// TIA Portal V19 export
FUNCTION_BLOCK "ALL_PUMPS"   // FB2, LAD
{ S7_Optimized_Access := 'TRUE' }
// stored: MemoryReserve 100, SetENOAutomatically false
   VAR
      PUMP_FB1_CP01 { S7_SetPoint := 'True'} : "PUMP_FB1";
      PUMP_FB1_AG01 { S7_SetPoint := 'True'} : "PUMP_FB1";
      PUMP_FB1_CHS_CP01 { S7_SetPoint := 'True'} : "PUMP_FB1";
      PUMP_FB1_CHS_CP02 { S7_SetPoint := 'True'} : "PUMP_FB1";
      PUMP_FB1_CHS_CP03 { S7_SetPoint := 'True'} : "PUMP_FB1";
      PUMP_FB1_R2_CP01 { S7_SetPoint := 'True'} : "PUMP_FB1";
      PUMP_FB1_R2_AG01 { S7_SetPoint := 'True'} : "PUMP_FB1";
      PUMP_FB1_R3_CP01 { S7_SetPoint := 'True'} : "PUMP_FB1";
      PUMP_FB1_R3_AG01 { S7_SetPoint := 'True'} : "PUMP_FB1";
      PUMP_FB1_R4_CP01 { S7_SetPoint := 'True'} : "PUMP_FB1";
      PUMP_FB1_R4_AG01 { S7_SetPoint := 'True'} : "PUMP_FB1";
      PUMP_FB1_R5_CP01 { S7_SetPoint := 'True'} : "PUMP_FB1";
      PUMP_FB1_R5_AG01 { S7_SetPoint := 'True'} : "PUMP_FB1";
      PUMP_FB1_R6_CP01 { S7_SetPoint := 'True'} : "PUMP_FB1";
      PUMP_FB1_R6_AG01 { S7_SetPoint := 'True'} : "PUMP_FB1";
      PUMP_FB1_R7_CP01 { S7_SetPoint := 'True'} : "PUMP_FB1";
      PUMP_FB1_R7_AG01 { S7_SetPoint := 'True'} : "PUMP_FB1";
      PUMP_FB1_R8_CP01 { S7_SetPoint := 'True'} : "PUMP_FB1";
      PUMP_FB1_R8_AG01 { S7_SetPoint := 'True'} : "PUMP_FB1";
      PUMP_FB1_R9_CP01 { S7_SetPoint := 'True'} : "PUMP_FB1";
      PUMP_FB1_R9_AG01 { S7_SetPoint := 'True'} : "PUMP_FB1";
      PUMP_FB1_R10_CP01 { S7_SetPoint := 'True'} : "PUMP_FB1";
      PUMP_FB1_R10_AG01 { S7_SetPoint := 'True'} : "PUMP_FB1";
      PUMP_FB1_R11_CP01 { S7_SetPoint := 'True'} : "PUMP_FB1";
      PUMP_FB1_R11_AG01 { S7_SetPoint := 'True'} : "PUMP_FB1";
      PUMP_FB1_R12_CP01 { S7_SetPoint := 'True'} : "PUMP_FB1";
      PUMP_FB1_R12_AG01 { S7_SetPoint := 'True'} : "PUMP_FB1";
      PUMP_FB1_R13_CP01 { S7_SetPoint := 'True'} : "PUMP_FB1";
      PUMP_FB1_R13_AG01 { S7_SetPoint := 'True'} : "PUMP_FB1";
      PUMP_FB1_R14_CP01 { S7_SetPoint := 'True'} : "PUMP_FB1";
      PUMP_FB1_R14_AG01 { S7_SetPoint := 'True'} : "PUMP_FB1";
      PUMP_FB1_R15_CP01 { S7_SetPoint := 'True'} : "PUMP_FB1";
      PUMP_FB1_R15_AG01 { S7_SetPoint := 'True'} : "PUMP_FB1";
      PUMP_FB1_R16_CP01 { S7_SetPoint := 'True'} : "PUMP_FB1";
      PUMP_FB1_R16_AG01 { S7_SetPoint := 'True'} : "PUMP_FB1";
      PUMP_FB1_R17_CP01 { S7_SetPoint := 'True'} : "PUMP_FB1";
      PUMP_FB1_R17_AG01 { S7_SetPoint := 'True'} : "PUMP_FB1";
      PUMP_FB1_R18_CP01 { S7_SetPoint := 'True'} : "PUMP_FB1";
      PUMP_FB1_R18_AG01 { S7_SetPoint := 'True'} : "PUMP_FB1";
      PUMP_FB1_CS_CP01 { S7_SetPoint := 'True'} : "PUMP_FB1";
      PUMP_FB1_CS_CP02 { S7_SetPoint := 'True'} : "PUMP_FB1";
      PUMP_FB1_CS_CP03 { S7_SetPoint := 'True'} : "PUMP_FB1";
      PUMP_FB1_UCHS_CP01 { S7_SetPoint := 'True'} : "PUMP_FB1";
      PUMP_FB1_UCHS_CP02 { S7_SetPoint := 'True'} : "PUMP_FB1";
      PUMP_FB1_UCHS_CP03 { S7_SetPoint := 'True'} : "PUMP_FB1";
      PUMP_FB1_HS_CP01 { S7_SetPoint := 'True'} : "PUMP_FB1";
      PUMP_FB1_HS_CP02 { S7_SetPoint := 'True'} : "PUMP_FB1";
      PUMP_FB1_HS_CP03 { S7_SetPoint := 'True'} : "PUMP_FB1";
      "PUMP_FB1_A/SCRB_001_CP01" { S7_SetPoint := 'True'} : "PUMP_FB1";
      "PUMP_FB1_A/SCRB_001_CP02" { S7_SetPoint := 'True'} : "PUMP_FB1";
      "PUMP_FB1_A/SCRB_002_CP01" { S7_SetPoint := 'True'} : "PUMP_FB1";
      "PUMP_FB1_A/SCRB_001_BL01" { S7_SetPoint := 'True'} : "PUMP_FB1";
      "PUMP_FB1_A/SCRB_002_BL02" { S7_SetPoint := 'True'} : "PUMP_FB1";
      "PUMP_FB1_AA/VP_01_CP01" { S7_SetPoint := 'True'} : "PUMP_FB1";
      "PUMP_FB1_A/VP_01_CP01" { S7_SetPoint := 'True'} : "PUMP_FB1";
   END_VAR
BEGIN

REGION Network 1: ***R1****
END_REGION

REGION Network 2: CP01
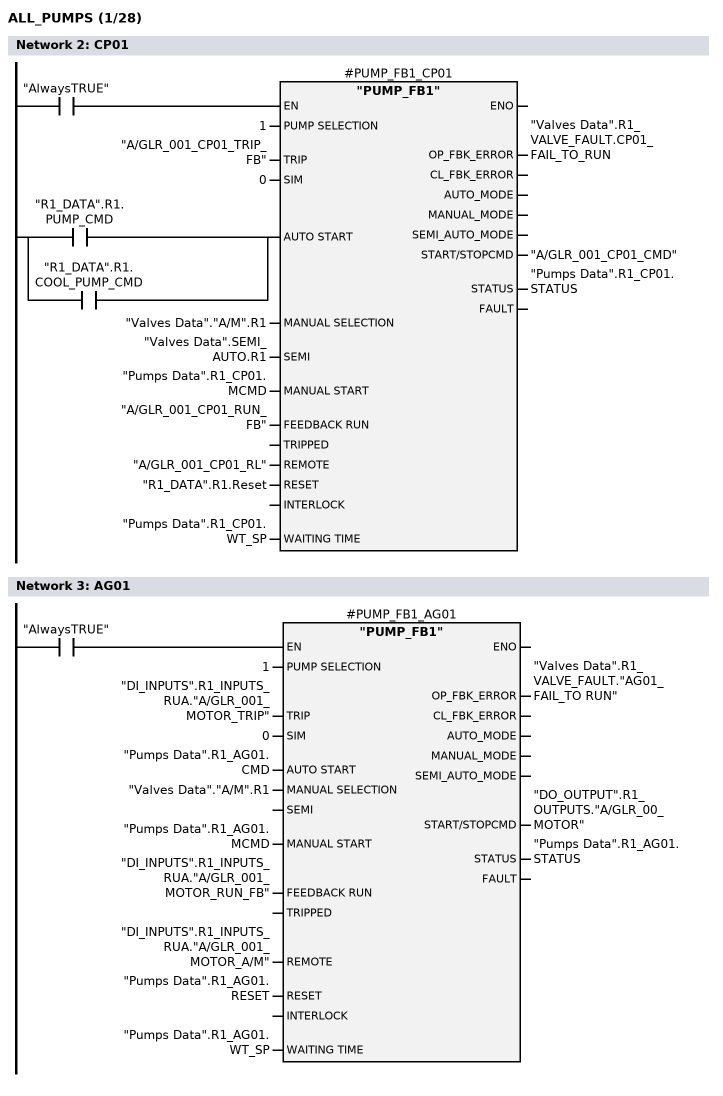
   RUNG wire#powerrail
      Contact( "AlwaysTRUE" )
      #PUMP_FB1_CP01("AUTO START" := wire#w1, "PUMP SELECTION" := 1, TRIP := "A/GLR_001_CP01_TRIP_FB", SIM := 0, "MANUAL SELECTION" := "Valves Data"."A/M".R1, SEMI := "Valves Data".SEMI_AUTO.R1, "MANUAL START" := "Pumps Data".R1_CP01.MCMD, "FEEDBACK RUN" := "A/GLR_001_CP01_RUN_FB", TRIPPED :=, REMOTE := "A/GLR_001_CP01_RL", RESET := "R1_DATA".R1.Reset, INTERLOCK :=, "WAITING TIME" := "Pumps Data".R1_CP01.WT_SP, OP_FBK_ERROR => "Valves Data".R1_VALVE_FAULT.CP01_FAIL_TO_RUN, CL_FBK_ERROR =>, AUTO_MODE =>, MANUAL_MODE =>, SEMI_AUTO_MODE =>, "START/STOPCMD" => "A/GLR_001_CP01_CMD", STATUS => "Pumps Data".R1_CP01.STATUS, FAULT =>)
   END_RUNG
   RUNG wire#powerrail
      Contact( "R1_DATA".R1.PUMP_CMD )
   END_RUNG wire#w1
   RUNG wire#powerrail
      Contact( "R1_DATA".R1.COOL_PUMP_CMD )
   END_RUNG wire#w1
   // the same network as SCL:
   IF "AlwaysTRUE" THEN
       #PUMP_FB1_CP01("PUMP SELECTION" := 1,   // "PUMP_FB1"
                      TRIP := "A/GLR_001_CP01_TRIP_FB",
                      SIM := 0,
                      "AUTO START" := "R1_DATA".R1.PUMP_CMD OR "R1_DATA".R1.COOL_PUMP_CMD,
                      "MANUAL SELECTION" := "Valves Data"."A/M".R1,
                      SEMI := "Valves Data".SEMI_AUTO.R1,
                      "MANUAL START" := "Pumps Data".R1_CP01.MCMD,
                      "FEEDBACK RUN" := "A/GLR_001_CP01_RUN_FB",
                      REMOTE := "A/GLR_001_CP01_RL",
                      RESET := "R1_DATA".R1.Reset,
                      "WAITING TIME" := "Pumps Data".R1_CP01.WT_SP,
                      OP_FBK_ERROR => "Valves Data".R1_VALVE_FAULT.CP01_FAIL_TO_RUN,
                      "START/STOPCMD" => "A/GLR_001_CP01_CMD",
                      STATUS => "Pumps Data".R1_CP01.STATUS);
   END_IF;
END_REGION

REGION Network 3: AG01
   RUNG wire#powerrail
      Contact( "AlwaysTRUE" )
      #PUMP_FB1_AG01("PUMP SELECTION" := 1, TRIP := "DI_INPUTS".R1_INPUTS_RUA."A/GLR_001_MOTOR_TRIP", SIM := 0, "AUTO START" := "Pumps Data".R1_AG01.CMD, "MANUAL SELECTION" := "Valves Data"."A/M".R1, SEMI :=, "MANUAL START" := "Pumps Data".R1_AG01.MCMD, "FEEDBACK RUN" := "DI_INPUTS".R1_INPUTS_RUA."A/GLR_001_MOTOR_RUN_FB", TRIPPED :=, REMOTE := "DI_INPUTS".R1_INPUTS_RUA."A/GLR_001_MOTOR_A/M", RESET := "Pumps Data".R1_AG01.RESET, INTERLOCK :=, "WAITING TIME" := "Pumps Data".R1_AG01.WT_SP, OP_FBK_ERROR => "Valves Data".R1_VALVE_FAULT."AG01_FAIL_TO RUN", CL_FBK_ERROR =>, AUTO_MODE =>, MANUAL_MODE =>, SEMI_AUTO_MODE =>, "START/STOPCMD" => "DO_OUTPUT".R1_OUTPUTS."A/GLR_00_MOTOR", STATUS => "Pumps Data".R1_AG01.STATUS, FAULT =>)
   END_RUNG
   // the same network as SCL:
   IF "AlwaysTRUE" THEN
       #PUMP_FB1_AG01("PUMP SELECTION" := 1,   // "PUMP_FB1"
                      TRIP := "DI_INPUTS".R1_INPUTS_RUA."A/GLR_001_MOTOR_TRIP",
                      SIM := 0,
                      "AUTO START" := "Pumps Data".R1_AG01.CMD,
                      "MANUAL SELECTION" := "Valves Data"."A/M".R1,
                      "MANUAL START" := "Pumps Data".R1_AG01.MCMD,
                      "FEEDBACK RUN" := "DI_INPUTS".R1_INPUTS_RUA."A/GLR_001_MOTOR_RUN_FB",
                      REMOTE := "DI_INPUTS".R1_INPUTS_RUA."A/GLR_001_MOTOR_A/M",
                      RESET := "Pumps Data".R1_AG01.RESET,
                      "WAITING TIME" := "Pumps Data".R1_AG01.WT_SP,
                      OP_FBK_ERROR => "Valves Data".R1_VALVE_FAULT."AG01_FAIL_TO RUN",
                      "START/STOPCMD" => "DO_OUTPUT".R1_OUTPUTS."A/GLR_00_MOTOR",
                      STATUS => "Pumps Data".R1_AG01.STATUS);
   END_IF;
END_REGION

REGION Network 4: CHS_CP01
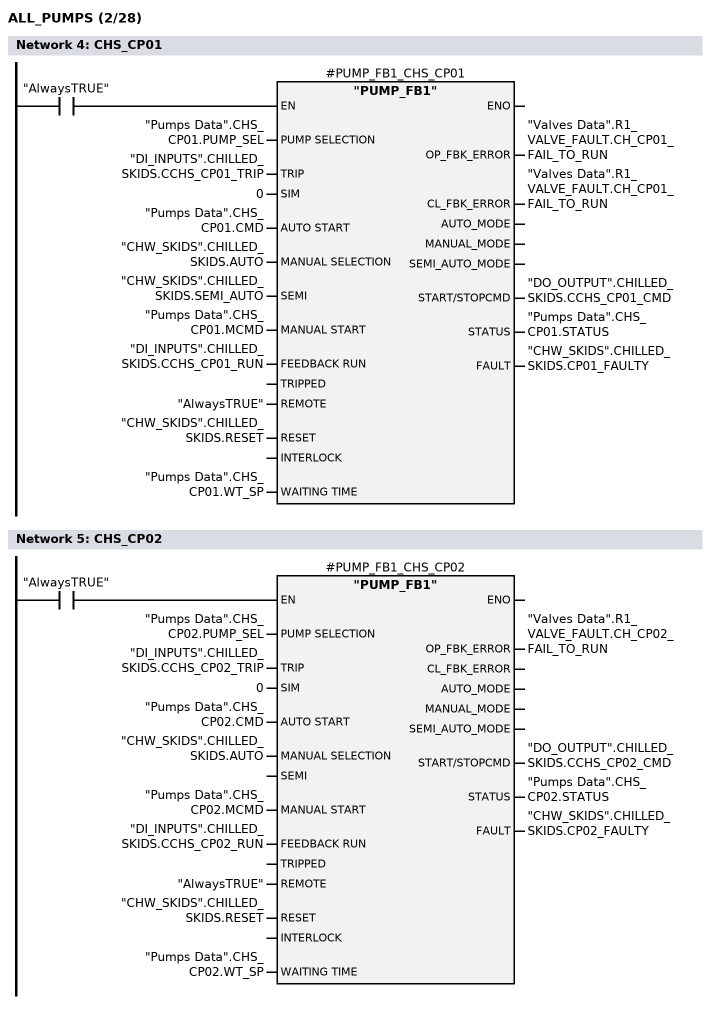
   RUNG wire#powerrail
      Contact( "AlwaysTRUE" )
      #PUMP_FB1_CHS_CP01("PUMP SELECTION" := "Pumps Data".CHS_CP01.PUMP_SEL, TRIP := "DI_INPUTS".CHILLED_SKIDS.CCHS_CP01_TRIP, SIM := 0, "AUTO START" := "Pumps Data".CHS_CP01.CMD, "MANUAL SELECTION" := "CHW_SKIDS".CHILLED_SKIDS.AUTO, SEMI := "CHW_SKIDS".CHILLED_SKIDS.SEMI_AUTO, "MANUAL START" := "Pumps Data".CHS_CP01.MCMD, "FEEDBACK RUN" := "DI_INPUTS".CHILLED_SKIDS.CCHS_CP01_RUN, TRIPPED :=, REMOTE := "AlwaysTRUE", RESET := "CHW_SKIDS".CHILLED_SKIDS.RESET, INTERLOCK :=, "WAITING TIME" := "Pumps Data".CHS_CP01.WT_SP, OP_FBK_ERROR => "Valves Data".R1_VALVE_FAULT.CH_CP01_FAIL_TO_RUN, CL_FBK_ERROR => "Valves Data".R1_VALVE_FAULT.CH_CP01_FAIL_TO_RUN, AUTO_MODE =>, MANUAL_MODE =>, SEMI_AUTO_MODE =>, "START/STOPCMD" => "DO_OUTPUT".CHILLED_SKIDS.CCHS_CP01_CMD, STATUS => "Pumps Data".CHS_CP01.STATUS, FAULT => "CHW_SKIDS".CHILLED_SKIDS.CP01_FAULTY)
   END_RUNG
   // the same network as SCL:
   IF "AlwaysTRUE" THEN
       #PUMP_FB1_CHS_CP01("PUMP SELECTION" := "Pumps Data".CHS_CP01.PUMP_SEL,   // "PUMP_FB1"
                          TRIP := "DI_INPUTS".CHILLED_SKIDS.CCHS_CP01_TRIP,
                          SIM := 0,
                          "AUTO START" := "Pumps Data".CHS_CP01.CMD,
                          "MANUAL SELECTION" := "CHW_SKIDS".CHILLED_SKIDS.AUTO,
                          SEMI := "CHW_SKIDS".CHILLED_SKIDS.SEMI_AUTO,
                          "MANUAL START" := "Pumps Data".CHS_CP01.MCMD,
                          "FEEDBACK RUN" := "DI_INPUTS".CHILLED_SKIDS.CCHS_CP01_RUN,
                          REMOTE := "AlwaysTRUE",
                          RESET := "CHW_SKIDS".CHILLED_SKIDS.RESET,
                          "WAITING TIME" := "Pumps Data".CHS_CP01.WT_SP,
                          OP_FBK_ERROR => "Valves Data".R1_VALVE_FAULT.CH_CP01_FAIL_TO_RUN,
                          CL_FBK_ERROR => "Valves Data".R1_VALVE_FAULT.CH_CP01_FAIL_TO_RUN,
                          "START/STOPCMD" => "DO_OUTPUT".CHILLED_SKIDS.CCHS_CP01_CMD,
                          STATUS => "Pumps Data".CHS_CP01.STATUS,
                          FAULT => "CHW_SKIDS".CHILLED_SKIDS.CP01_FAULTY);
   END_IF;
END_REGION

REGION Network 5: CHS_CP02
   RUNG wire#powerrail
      Contact( "AlwaysTRUE" )
      #PUMP_FB1_CHS_CP02("PUMP SELECTION" := "Pumps Data".CHS_CP02.PUMP_SEL, TRIP := "DI_INPUTS".CHILLED_SKIDS.CCHS_CP02_TRIP, SIM := 0, "AUTO START" := "Pumps Data".CHS_CP02.CMD, "MANUAL SELECTION" := "CHW_SKIDS".CHILLED_SKIDS.AUTO, SEMI :=, "MANUAL START" := "Pumps Data".CHS_CP02.MCMD, "FEEDBACK RUN" := "DI_INPUTS".CHILLED_SKIDS.CCHS_CP02_RUN, TRIPPED :=, REMOTE := "AlwaysTRUE", RESET := "CHW_SKIDS".CHILLED_SKIDS.RESET, INTERLOCK :=, "WAITING TIME" := "Pumps Data".CHS_CP02.WT_SP, OP_FBK_ERROR => "Valves Data".R1_VALVE_FAULT.CH_CP02_FAIL_TO_RUN, CL_FBK_ERROR =>, AUTO_MODE =>, MANUAL_MODE =>, SEMI_AUTO_MODE =>, "START/STOPCMD" => "DO_OUTPUT".CHILLED_SKIDS.CCHS_CP02_CMD, STATUS => "Pumps Data".CHS_CP02.STATUS, FAULT => "CHW_SKIDS".CHILLED_SKIDS.CP02_FAULTY)
   END_RUNG
   // the same network as SCL:
   IF "AlwaysTRUE" THEN
       #PUMP_FB1_CHS_CP02("PUMP SELECTION" := "Pumps Data".CHS_CP02.PUMP_SEL,   // "PUMP_FB1"
                          TRIP := "DI_INPUTS".CHILLED_SKIDS.CCHS_CP02_TRIP,
                          SIM := 0,
                          "AUTO START" := "Pumps Data".CHS_CP02.CMD,
                          "MANUAL SELECTION" := "CHW_SKIDS".CHILLED_SKIDS.AUTO,
                          "MANUAL START" := "Pumps Data".CHS_CP02.MCMD,
                          "FEEDBACK RUN" := "DI_INPUTS".CHILLED_SKIDS.CCHS_CP02_RUN,
                          REMOTE := "AlwaysTRUE",
                          RESET := "CHW_SKIDS".CHILLED_SKIDS.RESET,
                          "WAITING TIME" := "Pumps Data".CHS_CP02.WT_SP,
                          OP_FBK_ERROR => "Valves Data".R1_VALVE_FAULT.CH_CP02_FAIL_TO_RUN,
                          "START/STOPCMD" => "DO_OUTPUT".CHILLED_SKIDS.CCHS_CP02_CMD,
                          STATUS => "Pumps Data".CHS_CP02.STATUS,
                          FAULT => "CHW_SKIDS".CHILLED_SKIDS.CP02_FAULTY);
   END_IF;
END_REGION

REGION Network 6: CHS_CP03
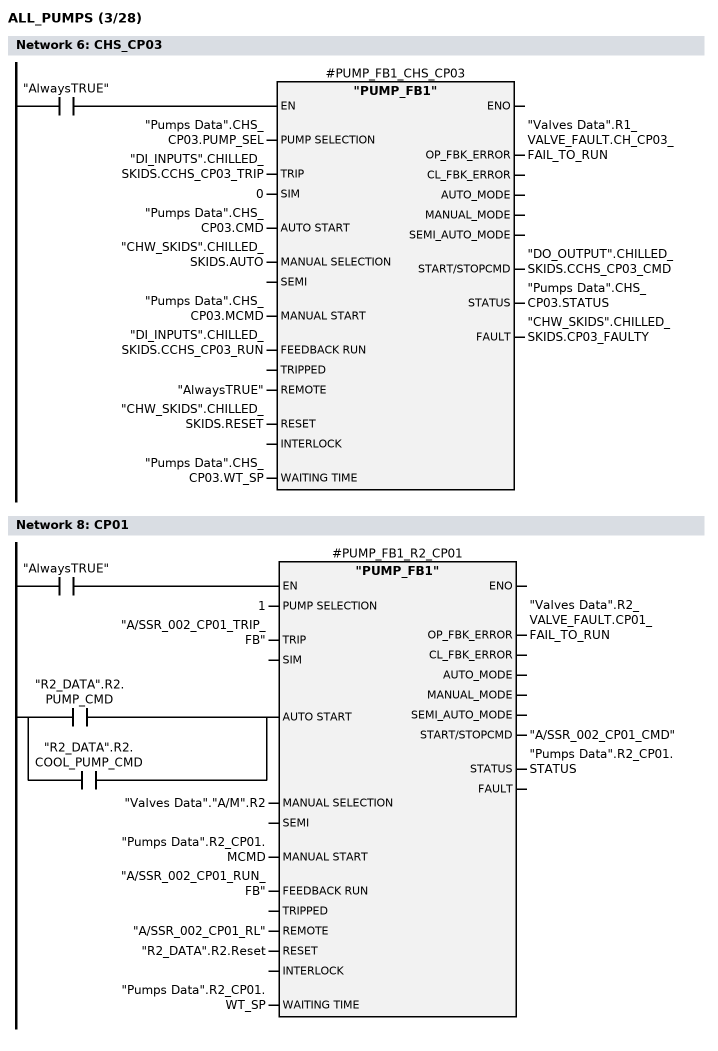
   RUNG wire#powerrail
      Contact( "AlwaysTRUE" )
      #PUMP_FB1_CHS_CP03("PUMP SELECTION" := "Pumps Data".CHS_CP03.PUMP_SEL, TRIP := "DI_INPUTS".CHILLED_SKIDS.CCHS_CP03_TRIP, SIM := 0, "AUTO START" := "Pumps Data".CHS_CP03.CMD, "MANUAL SELECTION" := "CHW_SKIDS".CHILLED_SKIDS.AUTO, SEMI :=, "MANUAL START" := "Pumps Data".CHS_CP03.MCMD, "FEEDBACK RUN" := "DI_INPUTS".CHILLED_SKIDS.CCHS_CP03_RUN, TRIPPED :=, REMOTE := "AlwaysTRUE", RESET := "CHW_SKIDS".CHILLED_SKIDS.RESET, INTERLOCK :=, "WAITING TIME" := "Pumps Data".CHS_CP03.WT_SP, OP_FBK_ERROR => "Valves Data".R1_VALVE_FAULT.CH_CP03_FAIL_TO_RUN, CL_FBK_ERROR =>, AUTO_MODE =>, MANUAL_MODE =>, SEMI_AUTO_MODE =>, "START/STOPCMD" => "DO_OUTPUT".CHILLED_SKIDS.CCHS_CP03_CMD, STATUS => "Pumps Data".CHS_CP03.STATUS, FAULT => "CHW_SKIDS".CHILLED_SKIDS.CP03_FAULTY)
   END_RUNG
   // the same network as SCL:
   IF "AlwaysTRUE" THEN
       #PUMP_FB1_CHS_CP03("PUMP SELECTION" := "Pumps Data".CHS_CP03.PUMP_SEL,   // "PUMP_FB1"
                          TRIP := "DI_INPUTS".CHILLED_SKIDS.CCHS_CP03_TRIP,
                          SIM := 0,
                          "AUTO START" := "Pumps Data".CHS_CP03.CMD,
                          "MANUAL SELECTION" := "CHW_SKIDS".CHILLED_SKIDS.AUTO,
                          "MANUAL START" := "Pumps Data".CHS_CP03.MCMD,
                          "FEEDBACK RUN" := "DI_INPUTS".CHILLED_SKIDS.CCHS_CP03_RUN,
                          REMOTE := "AlwaysTRUE",
                          RESET := "CHW_SKIDS".CHILLED_SKIDS.RESET,
                          "WAITING TIME" := "Pumps Data".CHS_CP03.WT_SP,
                          OP_FBK_ERROR => "Valves Data".R1_VALVE_FAULT.CH_CP03_FAIL_TO_RUN,
                          "START/STOPCMD" => "DO_OUTPUT".CHILLED_SKIDS.CCHS_CP03_CMD,
                          STATUS => "Pumps Data".CHS_CP03.STATUS,
                          FAULT => "CHW_SKIDS".CHILLED_SKIDS.CP03_FAULTY);
   END_IF;
END_REGION

REGION Network 7: ***R2****
END_REGION

REGION Network 8: CP01
   RUNG wire#powerrail
      Contact( "AlwaysTRUE" )
      #PUMP_FB1_R2_CP01("AUTO START" := wire#w1, "PUMP SELECTION" := 1, TRIP := "A/SSR_002_CP01_TRIP_FB", SIM :=, "MANUAL SELECTION" := "Valves Data"."A/M".R2, SEMI :=, "MANUAL START" := "Pumps Data".R2_CP01.MCMD, "FEEDBACK RUN" := "A/SSR_002_CP01_RUN_FB", TRIPPED :=, REMOTE := "A/SSR_002_CP01_RL", RESET := "R2_DATA".R2.Reset, INTERLOCK :=, "WAITING TIME" := "Pumps Data".R2_CP01.WT_SP, OP_FBK_ERROR => "Valves Data".R2_VALVE_FAULT.CP01_FAIL_TO_RUN, CL_FBK_ERROR =>, AUTO_MODE =>, MANUAL_MODE =>, SEMI_AUTO_MODE =>, "START/STOPCMD" => "A/SSR_002_CP01_CMD", STATUS => "Pumps Data".R2_CP01.STATUS, FAULT =>)
   END_RUNG
   RUNG wire#powerrail
      Contact( "R2_DATA".R2.PUMP_CMD )
   END_RUNG wire#w1
   RUNG wire#powerrail
      Contact( "R2_DATA".R2.COOL_PUMP_CMD )
   END_RUNG wire#w1
   // the same network as SCL:
   IF "AlwaysTRUE" THEN
       #PUMP_FB1_R2_CP01("PUMP SELECTION" := 1,   // "PUMP_FB1"
                         TRIP := "A/SSR_002_CP01_TRIP_FB",
                         "AUTO START" := "R2_DATA".R2.PUMP_CMD OR "R2_DATA".R2.COOL_PUMP_CMD,
                         "MANUAL SELECTION" := "Valves Data"."A/M".R2,
                         "MANUAL START" := "Pumps Data".R2_CP01.MCMD,
                         "FEEDBACK RUN" := "A/SSR_002_CP01_RUN_FB",
                         REMOTE := "A/SSR_002_CP01_RL",
                         RESET := "R2_DATA".R2.Reset,
                         "WAITING TIME" := "Pumps Data".R2_CP01.WT_SP,
                         OP_FBK_ERROR => "Valves Data".R2_VALVE_FAULT.CP01_FAIL_TO_RUN,
                         "START/STOPCMD" => "A/SSR_002_CP01_CMD",
                         STATUS => "Pumps Data".R2_CP01.STATUS);
   END_IF;
END_REGION

REGION Network 9: AG01
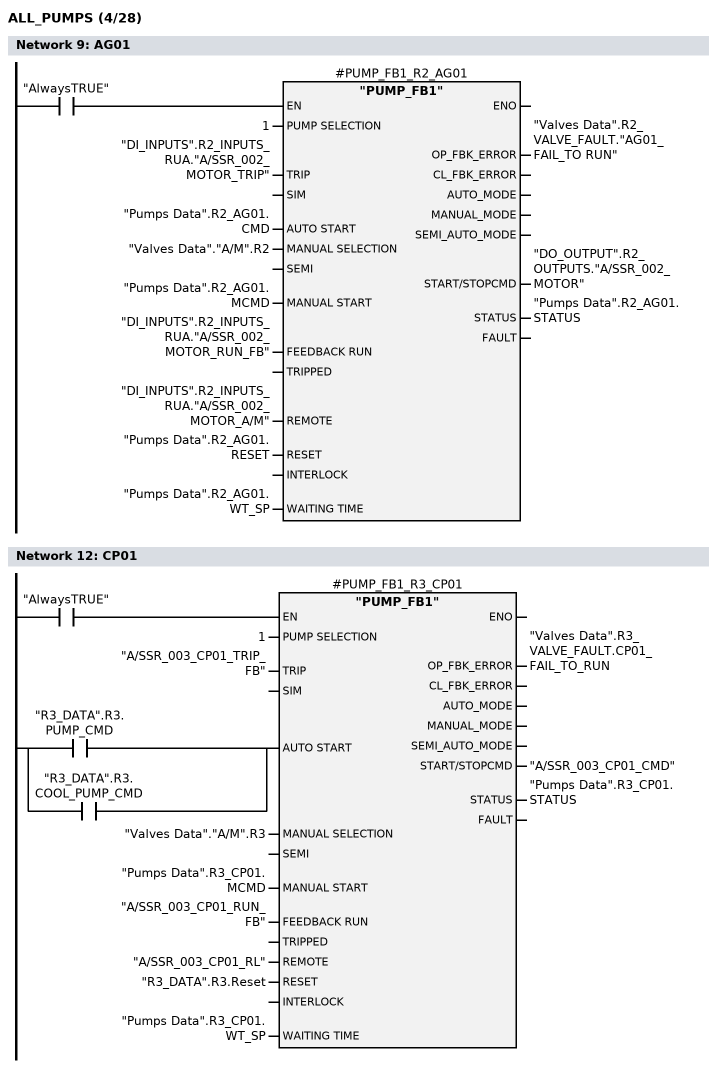
   RUNG wire#powerrail
      Contact( "AlwaysTRUE" )
      #PUMP_FB1_R2_AG01("PUMP SELECTION" := 1, TRIP := "DI_INPUTS".R2_INPUTS_RUA."A/SSR_002_MOTOR_TRIP", SIM :=, "AUTO START" := "Pumps Data".R2_AG01.CMD, "MANUAL SELECTION" := "Valves Data"."A/M".R2, SEMI :=, "MANUAL START" := "Pumps Data".R2_AG01.MCMD, "FEEDBACK RUN" := "DI_INPUTS".R2_INPUTS_RUA."A/SSR_002_MOTOR_RUN_FB", TRIPPED :=, REMOTE := "DI_INPUTS".R2_INPUTS_RUA."A/SSR_002_MOTOR_A/M", RESET := "Pumps Data".R2_AG01.RESET, INTERLOCK :=, "WAITING TIME" := "Pumps Data".R2_AG01.WT_SP, OP_FBK_ERROR => "Valves Data".R2_VALVE_FAULT."AG01_FAIL_TO RUN", CL_FBK_ERROR =>, AUTO_MODE =>, MANUAL_MODE =>, SEMI_AUTO_MODE =>, "START/STOPCMD" => "DO_OUTPUT".R2_OUTPUTS."A/SSR_002_MOTOR", STATUS => "Pumps Data".R2_AG01.STATUS, FAULT =>)
   END_RUNG
   // the same network as SCL:
   IF "AlwaysTRUE" THEN
       #PUMP_FB1_R2_AG01("PUMP SELECTION" := 1,   // "PUMP_FB1"
                         TRIP := "DI_INPUTS".R2_INPUTS_RUA."A/SSR_002_MOTOR_TRIP",
                         "AUTO START" := "Pumps Data".R2_AG01.CMD,
                         "MANUAL SELECTION" := "Valves Data"."A/M".R2,
                         "MANUAL START" := "Pumps Data".R2_AG01.MCMD,
                         "FEEDBACK RUN" := "DI_INPUTS".R2_INPUTS_RUA."A/SSR_002_MOTOR_RUN_FB",
                         REMOTE := "DI_INPUTS".R2_INPUTS_RUA."A/SSR_002_MOTOR_A/M",
                         RESET := "Pumps Data".R2_AG01.RESET,
                         "WAITING TIME" := "Pumps Data".R2_AG01.WT_SP,
                         OP_FBK_ERROR => "Valves Data".R2_VALVE_FAULT."AG01_FAIL_TO RUN",
                         "START/STOPCMD" => "DO_OUTPUT".R2_OUTPUTS."A/SSR_002_MOTOR",
                         STATUS => "Pumps Data".R2_AG01.STATUS);
   END_IF;
END_REGION

REGION Network 11: ***R3****
END_REGION

REGION Network 12: CP01
   RUNG wire#powerrail
      Contact( "AlwaysTRUE" )
      #PUMP_FB1_R3_CP01("AUTO START" := wire#w1, "PUMP SELECTION" := 1, TRIP := "A/SSR_003_CP01_TRIP_FB", SIM :=, "MANUAL SELECTION" := "Valves Data"."A/M".R3, SEMI :=, "MANUAL START" := "Pumps Data".R3_CP01.MCMD, "FEEDBACK RUN" := "A/SSR_003_CP01_RUN_FB", TRIPPED :=, REMOTE := "A/SSR_003_CP01_RL", RESET := "R3_DATA".R3.Reset, INTERLOCK :=, "WAITING TIME" := "Pumps Data".R3_CP01.WT_SP, OP_FBK_ERROR => "Valves Data".R3_VALVE_FAULT.CP01_FAIL_TO_RUN, CL_FBK_ERROR =>, AUTO_MODE =>, MANUAL_MODE =>, SEMI_AUTO_MODE =>, "START/STOPCMD" => "A/SSR_003_CP01_CMD", STATUS => "Pumps Data".R3_CP01.STATUS, FAULT =>)
   END_RUNG
   RUNG wire#powerrail
      Contact( "R3_DATA".R3.PUMP_CMD )
   END_RUNG wire#w1
   RUNG wire#powerrail
      Contact( "R3_DATA".R3.COOL_PUMP_CMD )
   END_RUNG wire#w1
   // the same network as SCL:
   IF "AlwaysTRUE" THEN
       #PUMP_FB1_R3_CP01("PUMP SELECTION" := 1,   // "PUMP_FB1"
                         TRIP := "A/SSR_003_CP01_TRIP_FB",
                         "AUTO START" := "R3_DATA".R3.PUMP_CMD OR "R3_DATA".R3.COOL_PUMP_CMD,
                         "MANUAL SELECTION" := "Valves Data"."A/M".R3,
                         "MANUAL START" := "Pumps Data".R3_CP01.MCMD,
                         "FEEDBACK RUN" := "A/SSR_003_CP01_RUN_FB",
                         REMOTE := "A/SSR_003_CP01_RL",
                         RESET := "R3_DATA".R3.Reset,
                         "WAITING TIME" := "Pumps Data".R3_CP01.WT_SP,
                         OP_FBK_ERROR => "Valves Data".R3_VALVE_FAULT.CP01_FAIL_TO_RUN,
                         "START/STOPCMD" => "A/SSR_003_CP01_CMD",
                         STATUS => "Pumps Data".R3_CP01.STATUS);
   END_IF;
END_REGION

REGION Network 13: AG01
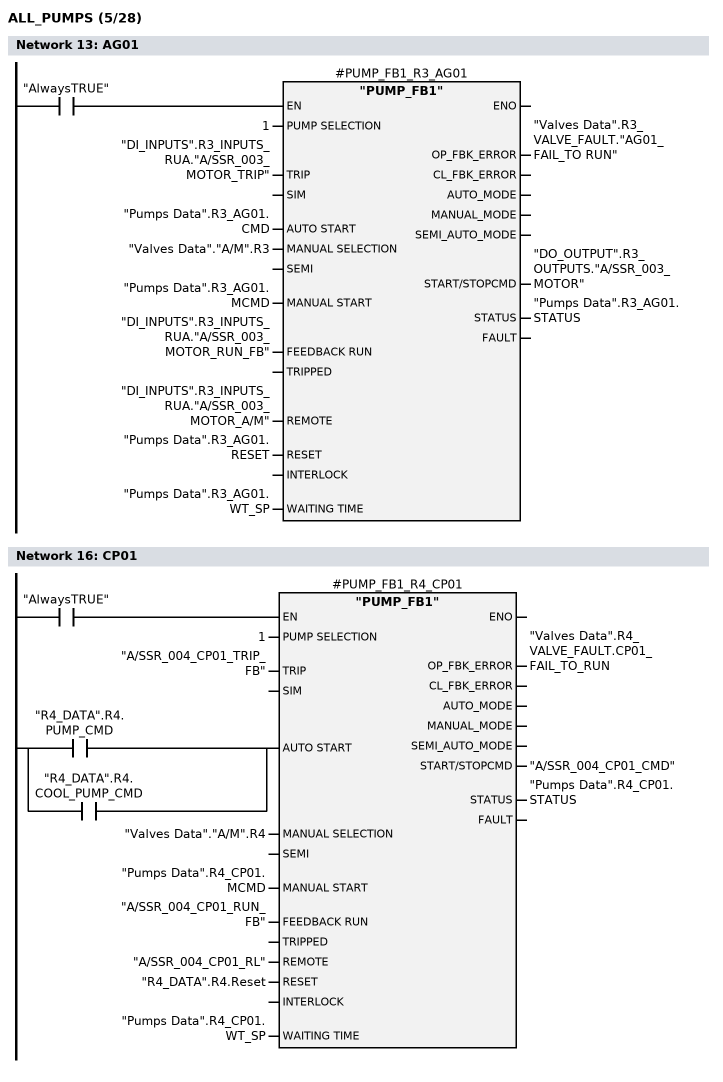
   RUNG wire#powerrail
      Contact( "AlwaysTRUE" )
      #PUMP_FB1_R3_AG01("PUMP SELECTION" := 1, TRIP := "DI_INPUTS".R3_INPUTS_RUA."A/SSR_003_MOTOR_TRIP", SIM :=, "AUTO START" := "Pumps Data".R3_AG01.CMD, "MANUAL SELECTION" := "Valves Data"."A/M".R3, SEMI :=, "MANUAL START" := "Pumps Data".R3_AG01.MCMD, "FEEDBACK RUN" := "DI_INPUTS".R3_INPUTS_RUA."A/SSR_003_MOTOR_RUN_FB", TRIPPED :=, REMOTE := "DI_INPUTS".R3_INPUTS_RUA."A/SSR_003_MOTOR_A/M", RESET := "Pumps Data".R3_AG01.RESET, INTERLOCK :=, "WAITING TIME" := "Pumps Data".R3_AG01.WT_SP, OP_FBK_ERROR => "Valves Data".R3_VALVE_FAULT."AG01_FAIL_TO RUN", CL_FBK_ERROR =>, AUTO_MODE =>, MANUAL_MODE =>, SEMI_AUTO_MODE =>, "START/STOPCMD" => "DO_OUTPUT".R3_OUTPUTS."A/SSR_003_MOTOR", STATUS => "Pumps Data".R3_AG01.STATUS, FAULT =>)
   END_RUNG
   // the same network as SCL:
   IF "AlwaysTRUE" THEN
       #PUMP_FB1_R3_AG01("PUMP SELECTION" := 1,   // "PUMP_FB1"
                         TRIP := "DI_INPUTS".R3_INPUTS_RUA."A/SSR_003_MOTOR_TRIP",
                         "AUTO START" := "Pumps Data".R3_AG01.CMD,
                         "MANUAL SELECTION" := "Valves Data"."A/M".R3,
                         "MANUAL START" := "Pumps Data".R3_AG01.MCMD,
                         "FEEDBACK RUN" := "DI_INPUTS".R3_INPUTS_RUA."A/SSR_003_MOTOR_RUN_FB",
                         REMOTE := "DI_INPUTS".R3_INPUTS_RUA."A/SSR_003_MOTOR_A/M",
                         RESET := "Pumps Data".R3_AG01.RESET,
                         "WAITING TIME" := "Pumps Data".R3_AG01.WT_SP,
                         OP_FBK_ERROR => "Valves Data".R3_VALVE_FAULT."AG01_FAIL_TO RUN",
                         "START/STOPCMD" => "DO_OUTPUT".R3_OUTPUTS."A/SSR_003_MOTOR",
                         STATUS => "Pumps Data".R3_AG01.STATUS);
   END_IF;
END_REGION

REGION Network 15: ***R4****
END_REGION

REGION Network 16: CP01
   RUNG wire#powerrail
      Contact( "AlwaysTRUE" )
      #PUMP_FB1_R4_CP01("AUTO START" := wire#w1, "PUMP SELECTION" := 1, TRIP := "A/SSR_004_CP01_TRIP_FB", SIM :=, "MANUAL SELECTION" := "Valves Data"."A/M".R4, SEMI :=, "MANUAL START" := "Pumps Data".R4_CP01.MCMD, "FEEDBACK RUN" := "A/SSR_004_CP01_RUN_FB", TRIPPED :=, REMOTE := "A/SSR_004_CP01_RL", RESET := "R4_DATA".R4.Reset, INTERLOCK :=, "WAITING TIME" := "Pumps Data".R4_CP01.WT_SP, OP_FBK_ERROR => "Valves Data".R4_VALVE_FAULT.CP01_FAIL_TO_RUN, CL_FBK_ERROR =>, AUTO_MODE =>, MANUAL_MODE =>, SEMI_AUTO_MODE =>, "START/STOPCMD" => "A/SSR_004_CP01_CMD", STATUS => "Pumps Data".R4_CP01.STATUS, FAULT =>)
   END_RUNG
   RUNG wire#powerrail
      Contact( "R4_DATA".R4.PUMP_CMD )
   END_RUNG wire#w1
   RUNG wire#powerrail
      Contact( "R4_DATA".R4.COOL_PUMP_CMD )
   END_RUNG wire#w1
   // the same network as SCL:
   IF "AlwaysTRUE" THEN
       #PUMP_FB1_R4_CP01("PUMP SELECTION" := 1,   // "PUMP_FB1"
                         TRIP := "A/SSR_004_CP01_TRIP_FB",
                         "AUTO START" := "R4_DATA".R4.PUMP_CMD OR "R4_DATA".R4.COOL_PUMP_CMD,
                         "MANUAL SELECTION" := "Valves Data"."A/M".R4,
                         "MANUAL START" := "Pumps Data".R4_CP01.MCMD,
                         "FEEDBACK RUN" := "A/SSR_004_CP01_RUN_FB",
                         REMOTE := "A/SSR_004_CP01_RL",
                         RESET := "R4_DATA".R4.Reset,
                         "WAITING TIME" := "Pumps Data".R4_CP01.WT_SP,
                         OP_FBK_ERROR => "Valves Data".R4_VALVE_FAULT.CP01_FAIL_TO_RUN,
                         "START/STOPCMD" => "A/SSR_004_CP01_CMD",
                         STATUS => "Pumps Data".R4_CP01.STATUS);
   END_IF;
END_REGION

REGION Network 17: AG01
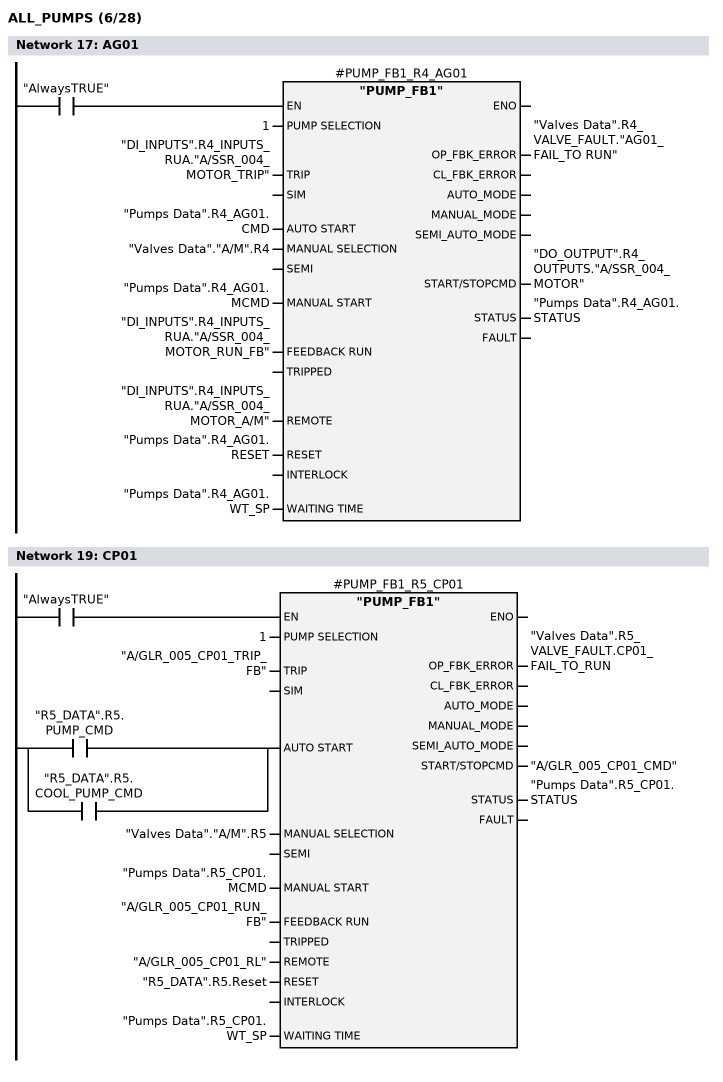
   RUNG wire#powerrail
      Contact( "AlwaysTRUE" )
      #PUMP_FB1_R4_AG01("PUMP SELECTION" := 1, TRIP := "DI_INPUTS".R4_INPUTS_RUA."A/SSR_004_MOTOR_TRIP", SIM :=, "AUTO START" := "Pumps Data".R4_AG01.CMD, "MANUAL SELECTION" := "Valves Data"."A/M".R4, SEMI :=, "MANUAL START" := "Pumps Data".R4_AG01.MCMD, "FEEDBACK RUN" := "DI_INPUTS".R4_INPUTS_RUA."A/SSR_004_MOTOR_RUN_FB", TRIPPED :=, REMOTE := "DI_INPUTS".R4_INPUTS_RUA."A/SSR_004_MOTOR_A/M", RESET := "Pumps Data".R4_AG01.RESET, INTERLOCK :=, "WAITING TIME" := "Pumps Data".R4_AG01.WT_SP, OP_FBK_ERROR => "Valves Data".R4_VALVE_FAULT."AG01_FAIL_TO RUN", CL_FBK_ERROR =>, AUTO_MODE =>, MANUAL_MODE =>, SEMI_AUTO_MODE =>, "START/STOPCMD" => "DO_OUTPUT".R4_OUTPUTS."A/SSR_004_MOTOR", STATUS => "Pumps Data".R4_AG01.STATUS, FAULT =>)
   END_RUNG
   // the same network as SCL:
   IF "AlwaysTRUE" THEN
       #PUMP_FB1_R4_AG01("PUMP SELECTION" := 1,   // "PUMP_FB1"
                         TRIP := "DI_INPUTS".R4_INPUTS_RUA."A/SSR_004_MOTOR_TRIP",
                         "AUTO START" := "Pumps Data".R4_AG01.CMD,
                         "MANUAL SELECTION" := "Valves Data"."A/M".R4,
                         "MANUAL START" := "Pumps Data".R4_AG01.MCMD,
                         "FEEDBACK RUN" := "DI_INPUTS".R4_INPUTS_RUA."A/SSR_004_MOTOR_RUN_FB",
                         REMOTE := "DI_INPUTS".R4_INPUTS_RUA."A/SSR_004_MOTOR_A/M",
                         RESET := "Pumps Data".R4_AG01.RESET,
                         "WAITING TIME" := "Pumps Data".R4_AG01.WT_SP,
                         OP_FBK_ERROR => "Valves Data".R4_VALVE_FAULT."AG01_FAIL_TO RUN",
                         "START/STOPCMD" => "DO_OUTPUT".R4_OUTPUTS."A/SSR_004_MOTOR",
                         STATUS => "Pumps Data".R4_AG01.STATUS);
   END_IF;
END_REGION

REGION Network 18: ***R5****
END_REGION

REGION Network 19: CP01
   RUNG wire#powerrail
      Contact( "AlwaysTRUE" )
      #PUMP_FB1_R5_CP01("AUTO START" := wire#w1, "PUMP SELECTION" := 1, TRIP := "A/GLR_005_CP01_TRIP_FB", SIM :=, "MANUAL SELECTION" := "Valves Data"."A/M".R5, SEMI :=, "MANUAL START" := "Pumps Data".R5_CP01.MCMD, "FEEDBACK RUN" := "A/GLR_005_CP01_RUN_FB", TRIPPED :=, REMOTE := "A/GLR_005_CP01_RL", RESET := "R5_DATA".R5.Reset, INTERLOCK :=, "WAITING TIME" := "Pumps Data".R5_CP01.WT_SP, OP_FBK_ERROR => "Valves Data".R5_VALVE_FAULT.CP01_FAIL_TO_RUN, CL_FBK_ERROR =>, AUTO_MODE =>, MANUAL_MODE =>, SEMI_AUTO_MODE =>, "START/STOPCMD" => "A/GLR_005_CP01_CMD", STATUS => "Pumps Data".R5_CP01.STATUS, FAULT =>)
   END_RUNG
   RUNG wire#powerrail
      Contact( "R5_DATA".R5.PUMP_CMD )
   END_RUNG wire#w1
   RUNG wire#powerrail
      Contact( "R5_DATA".R5.COOL_PUMP_CMD )
   END_RUNG wire#w1
   // the same network as SCL:
   IF "AlwaysTRUE" THEN
       #PUMP_FB1_R5_CP01("PUMP SELECTION" := 1,   // "PUMP_FB1"
                         TRIP := "A/GLR_005_CP01_TRIP_FB",
                         "AUTO START" := "R5_DATA".R5.PUMP_CMD OR "R5_DATA".R5.COOL_PUMP_CMD,
                         "MANUAL SELECTION" := "Valves Data"."A/M".R5,
                         "MANUAL START" := "Pumps Data".R5_CP01.MCMD,
                         "FEEDBACK RUN" := "A/GLR_005_CP01_RUN_FB",
                         REMOTE := "A/GLR_005_CP01_RL",
                         RESET := "R5_DATA".R5.Reset,
                         "WAITING TIME" := "Pumps Data".R5_CP01.WT_SP,
                         OP_FBK_ERROR => "Valves Data".R5_VALVE_FAULT.CP01_FAIL_TO_RUN,
                         "START/STOPCMD" => "A/GLR_005_CP01_CMD",
                         STATUS => "Pumps Data".R5_CP01.STATUS);
   END_IF;
END_REGION

REGION Network 20: AG01
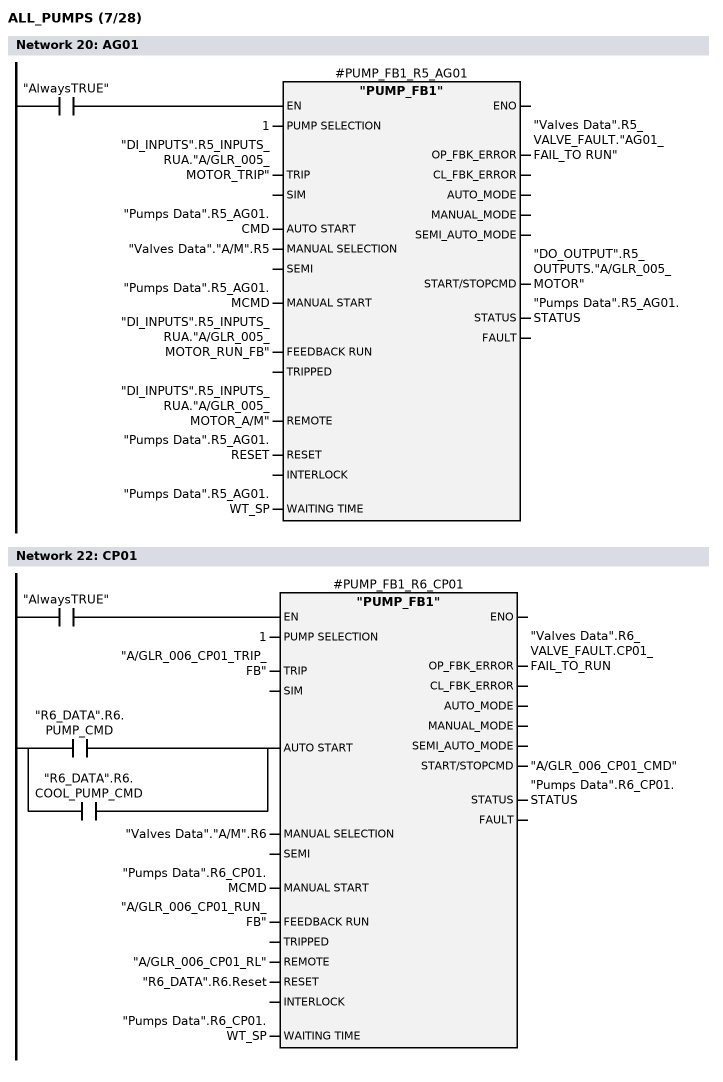
   RUNG wire#powerrail
      Contact( "AlwaysTRUE" )
      #PUMP_FB1_R5_AG01("PUMP SELECTION" := 1, TRIP := "DI_INPUTS".R5_INPUTS_RUA."A/GLR_005_MOTOR_TRIP", SIM :=, "AUTO START" := "Pumps Data".R5_AG01.CMD, "MANUAL SELECTION" := "Valves Data"."A/M".R5, SEMI :=, "MANUAL START" := "Pumps Data".R5_AG01.MCMD, "FEEDBACK RUN" := "DI_INPUTS".R5_INPUTS_RUA."A/GLR_005_MOTOR_RUN_FB", TRIPPED :=, REMOTE := "DI_INPUTS".R5_INPUTS_RUA."A/GLR_005_MOTOR_A/M", RESET := "Pumps Data".R5_AG01.RESET, INTERLOCK :=, "WAITING TIME" := "Pumps Data".R5_AG01.WT_SP, OP_FBK_ERROR => "Valves Data".R5_VALVE_FAULT."AG01_FAIL_TO RUN", CL_FBK_ERROR =>, AUTO_MODE =>, MANUAL_MODE =>, SEMI_AUTO_MODE =>, "START/STOPCMD" => "DO_OUTPUT".R5_OUTPUTS."A/GLR_005_MOTOR", STATUS => "Pumps Data".R5_AG01.STATUS, FAULT =>)
   END_RUNG
   // the same network as SCL:
   IF "AlwaysTRUE" THEN
       #PUMP_FB1_R5_AG01("PUMP SELECTION" := 1,   // "PUMP_FB1"
                         TRIP := "DI_INPUTS".R5_INPUTS_RUA."A/GLR_005_MOTOR_TRIP",
                         "AUTO START" := "Pumps Data".R5_AG01.CMD,
                         "MANUAL SELECTION" := "Valves Data"."A/M".R5,
                         "MANUAL START" := "Pumps Data".R5_AG01.MCMD,
                         "FEEDBACK RUN" := "DI_INPUTS".R5_INPUTS_RUA."A/GLR_005_MOTOR_RUN_FB",
                         REMOTE := "DI_INPUTS".R5_INPUTS_RUA."A/GLR_005_MOTOR_A/M",
                         RESET := "Pumps Data".R5_AG01.RESET,
                         "WAITING TIME" := "Pumps Data".R5_AG01.WT_SP,
                         OP_FBK_ERROR => "Valves Data".R5_VALVE_FAULT."AG01_FAIL_TO RUN",
                         "START/STOPCMD" => "DO_OUTPUT".R5_OUTPUTS."A/GLR_005_MOTOR",
                         STATUS => "Pumps Data".R5_AG01.STATUS);
   END_IF;
END_REGION

REGION Network 21: ***R6****
END_REGION

REGION Network 22: CP01
   RUNG wire#powerrail
      Contact( "AlwaysTRUE" )
      #PUMP_FB1_R6_CP01("AUTO START" := wire#w1, "PUMP SELECTION" := 1, TRIP := "A/GLR_006_CP01_TRIP_FB", SIM :=, "MANUAL SELECTION" := "Valves Data"."A/M".R6, SEMI :=, "MANUAL START" := "Pumps Data".R6_CP01.MCMD, "FEEDBACK RUN" := "A/GLR_006_CP01_RUN_FB", TRIPPED :=, REMOTE := "A/GLR_006_CP01_RL", RESET := "R6_DATA".R6.Reset, INTERLOCK :=, "WAITING TIME" := "Pumps Data".R6_CP01.WT_SP, OP_FBK_ERROR => "Valves Data".R6_VALVE_FAULT.CP01_FAIL_TO_RUN, CL_FBK_ERROR =>, AUTO_MODE =>, MANUAL_MODE =>, SEMI_AUTO_MODE =>, "START/STOPCMD" => "A/GLR_006_CP01_CMD", STATUS => "Pumps Data".R6_CP01.STATUS, FAULT =>)
   END_RUNG
   RUNG wire#powerrail
      Contact( "R6_DATA".R6.PUMP_CMD )
   END_RUNG wire#w1
   RUNG wire#powerrail
      Contact( "R6_DATA".R6.COOL_PUMP_CMD )
   END_RUNG wire#w1
   // the same network as SCL:
   IF "AlwaysTRUE" THEN
       #PUMP_FB1_R6_CP01("PUMP SELECTION" := 1,   // "PUMP_FB1"
                         TRIP := "A/GLR_006_CP01_TRIP_FB",
                         "AUTO START" := "R6_DATA".R6.PUMP_CMD OR "R6_DATA".R6.COOL_PUMP_CMD,
                         "MANUAL SELECTION" := "Valves Data"."A/M".R6,
                         "MANUAL START" := "Pumps Data".R6_CP01.MCMD,
                         "FEEDBACK RUN" := "A/GLR_006_CP01_RUN_FB",
                         REMOTE := "A/GLR_006_CP01_RL",
                         RESET := "R6_DATA".R6.Reset,
                         "WAITING TIME" := "Pumps Data".R6_CP01.WT_SP,
                         OP_FBK_ERROR => "Valves Data".R6_VALVE_FAULT.CP01_FAIL_TO_RUN,
                         "START/STOPCMD" => "A/GLR_006_CP01_CMD",
                         STATUS => "Pumps Data".R6_CP01.STATUS);
   END_IF;
END_REGION

REGION Network 23: AG01
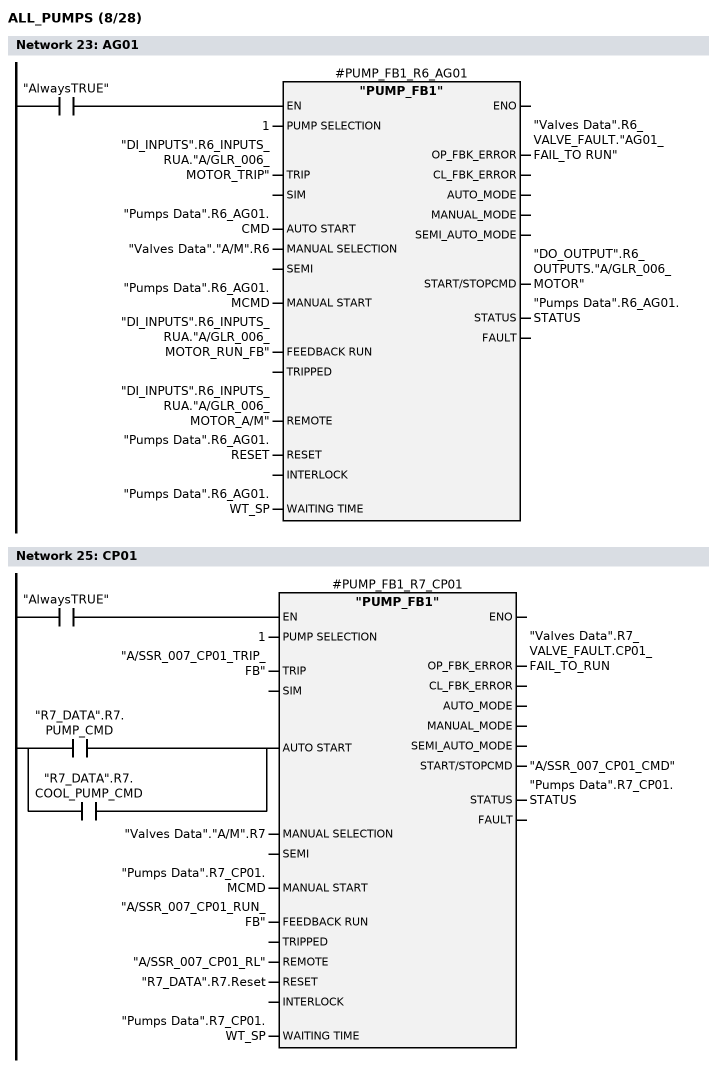
   RUNG wire#powerrail
      Contact( "AlwaysTRUE" )
      #PUMP_FB1_R6_AG01("PUMP SELECTION" := 1, TRIP := "DI_INPUTS".R6_INPUTS_RUA."A/GLR_006_MOTOR_TRIP", SIM :=, "AUTO START" := "Pumps Data".R6_AG01.CMD, "MANUAL SELECTION" := "Valves Data"."A/M".R6, SEMI :=, "MANUAL START" := "Pumps Data".R6_AG01.MCMD, "FEEDBACK RUN" := "DI_INPUTS".R6_INPUTS_RUA."A/GLR_006_MOTOR_RUN_FB", TRIPPED :=, REMOTE := "DI_INPUTS".R6_INPUTS_RUA."A/GLR_006_MOTOR_A/M", RESET := "Pumps Data".R6_AG01.RESET, INTERLOCK :=, "WAITING TIME" := "Pumps Data".R6_AG01.WT_SP, OP_FBK_ERROR => "Valves Data".R6_VALVE_FAULT."AG01_FAIL_TO RUN", CL_FBK_ERROR =>, AUTO_MODE =>, MANUAL_MODE =>, SEMI_AUTO_MODE =>, "START/STOPCMD" => "DO_OUTPUT".R6_OUTPUTS."A/GLR_006_MOTOR", STATUS => "Pumps Data".R6_AG01.STATUS, FAULT =>)
   END_RUNG
   // the same network as SCL:
   IF "AlwaysTRUE" THEN
       #PUMP_FB1_R6_AG01("PUMP SELECTION" := 1,   // "PUMP_FB1"
                         TRIP := "DI_INPUTS".R6_INPUTS_RUA."A/GLR_006_MOTOR_TRIP",
                         "AUTO START" := "Pumps Data".R6_AG01.CMD,
                         "MANUAL SELECTION" := "Valves Data"."A/M".R6,
                         "MANUAL START" := "Pumps Data".R6_AG01.MCMD,
                         "FEEDBACK RUN" := "DI_INPUTS".R6_INPUTS_RUA."A/GLR_006_MOTOR_RUN_FB",
                         REMOTE := "DI_INPUTS".R6_INPUTS_RUA."A/GLR_006_MOTOR_A/M",
                         RESET := "Pumps Data".R6_AG01.RESET,
                         "WAITING TIME" := "Pumps Data".R6_AG01.WT_SP,
                         OP_FBK_ERROR => "Valves Data".R6_VALVE_FAULT."AG01_FAIL_TO RUN",
                         "START/STOPCMD" => "DO_OUTPUT".R6_OUTPUTS."A/GLR_006_MOTOR",
                         STATUS => "Pumps Data".R6_AG01.STATUS);
   END_IF;
END_REGION

REGION Network 24: ***R7****
END_REGION

REGION Network 25: CP01
   RUNG wire#powerrail
      Contact( "AlwaysTRUE" )
      #PUMP_FB1_R7_CP01("AUTO START" := wire#w1, "PUMP SELECTION" := 1, TRIP := "A/SSR_007_CP01_TRIP_FB", SIM :=, "MANUAL SELECTION" := "Valves Data"."A/M".R7, SEMI :=, "MANUAL START" := "Pumps Data".R7_CP01.MCMD, "FEEDBACK RUN" := "A/SSR_007_CP01_RUN_FB", TRIPPED :=, REMOTE := "A/SSR_007_CP01_RL", RESET := "R7_DATA".R7.Reset, INTERLOCK :=, "WAITING TIME" := "Pumps Data".R7_CP01.WT_SP, OP_FBK_ERROR => "Valves Data".R7_VALVE_FAULT.CP01_FAIL_TO_RUN, CL_FBK_ERROR =>, AUTO_MODE =>, MANUAL_MODE =>, SEMI_AUTO_MODE =>, "START/STOPCMD" => "A/SSR_007_CP01_CMD", STATUS => "Pumps Data".R7_CP01.STATUS, FAULT =>)
   END_RUNG
   RUNG wire#powerrail
      Contact( "R7_DATA".R7.PUMP_CMD )
   END_RUNG wire#w1
   RUNG wire#powerrail
      Contact( "R7_DATA".R7.COOL_PUMP_CMD )
   END_RUNG wire#w1
   // the same network as SCL:
   IF "AlwaysTRUE" THEN
       #PUMP_FB1_R7_CP01("PUMP SELECTION" := 1,   // "PUMP_FB1"
                         TRIP := "A/SSR_007_CP01_TRIP_FB",
                         "AUTO START" := "R7_DATA".R7.PUMP_CMD OR "R7_DATA".R7.COOL_PUMP_CMD,
                         "MANUAL SELECTION" := "Valves Data"."A/M".R7,
                         "MANUAL START" := "Pumps Data".R7_CP01.MCMD,
                         "FEEDBACK RUN" := "A/SSR_007_CP01_RUN_FB",
                         REMOTE := "A/SSR_007_CP01_RL",
                         RESET := "R7_DATA".R7.Reset,
                         "WAITING TIME" := "Pumps Data".R7_CP01.WT_SP,
                         OP_FBK_ERROR => "Valves Data".R7_VALVE_FAULT.CP01_FAIL_TO_RUN,
                         "START/STOPCMD" => "A/SSR_007_CP01_CMD",
                         STATUS => "Pumps Data".R7_CP01.STATUS);
   END_IF;
END_REGION

REGION Network 26: AG01
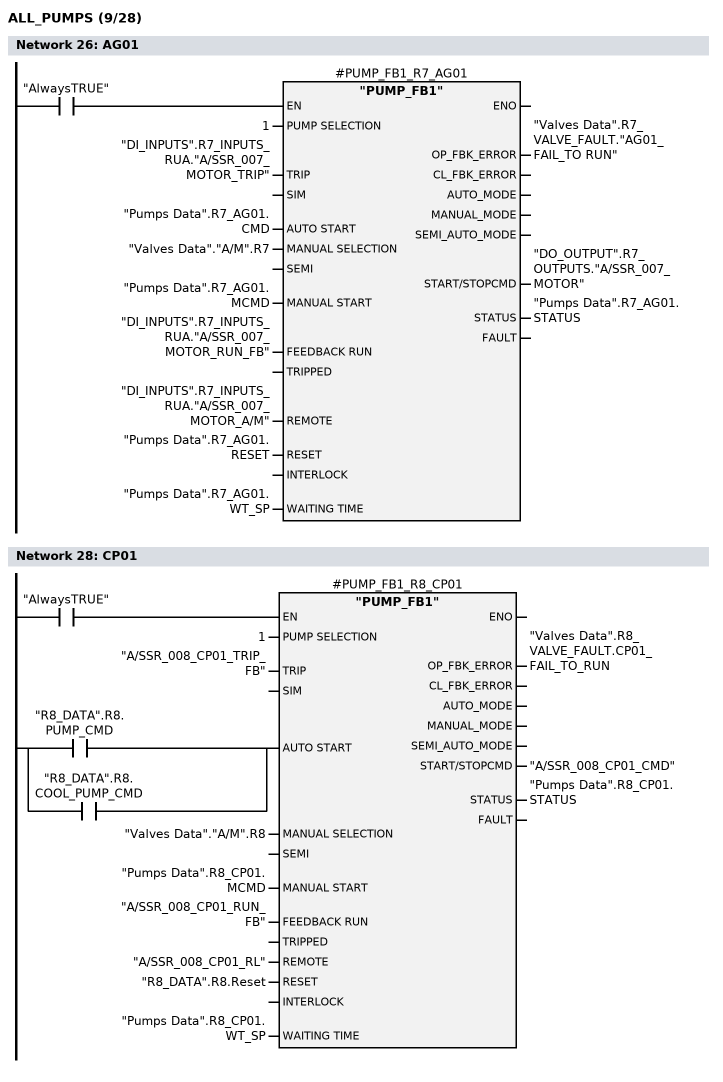
   RUNG wire#powerrail
      Contact( "AlwaysTRUE" )
      #PUMP_FB1_R7_AG01("PUMP SELECTION" := 1, TRIP := "DI_INPUTS".R7_INPUTS_RUA."A/SSR_007_MOTOR_TRIP", SIM :=, "AUTO START" := "Pumps Data".R7_AG01.CMD, "MANUAL SELECTION" := "Valves Data"."A/M".R7, SEMI :=, "MANUAL START" := "Pumps Data".R7_AG01.MCMD, "FEEDBACK RUN" := "DI_INPUTS".R7_INPUTS_RUA."A/SSR_007_MOTOR_RUN_FB", TRIPPED :=, REMOTE := "DI_INPUTS".R7_INPUTS_RUA."A/SSR_007_MOTOR_A/M", RESET := "Pumps Data".R7_AG01.RESET, INTERLOCK :=, "WAITING TIME" := "Pumps Data".R7_AG01.WT_SP, OP_FBK_ERROR => "Valves Data".R7_VALVE_FAULT."AG01_FAIL_TO RUN", CL_FBK_ERROR =>, AUTO_MODE =>, MANUAL_MODE =>, SEMI_AUTO_MODE =>, "START/STOPCMD" => "DO_OUTPUT".R7_OUTPUTS."A/SSR_007_MOTOR", STATUS => "Pumps Data".R7_AG01.STATUS, FAULT =>)
   END_RUNG
   // the same network as SCL:
   IF "AlwaysTRUE" THEN
       #PUMP_FB1_R7_AG01("PUMP SELECTION" := 1,   // "PUMP_FB1"
                         TRIP := "DI_INPUTS".R7_INPUTS_RUA."A/SSR_007_MOTOR_TRIP",
                         "AUTO START" := "Pumps Data".R7_AG01.CMD,
                         "MANUAL SELECTION" := "Valves Data"."A/M".R7,
                         "MANUAL START" := "Pumps Data".R7_AG01.MCMD,
                         "FEEDBACK RUN" := "DI_INPUTS".R7_INPUTS_RUA."A/SSR_007_MOTOR_RUN_FB",
                         REMOTE := "DI_INPUTS".R7_INPUTS_RUA."A/SSR_007_MOTOR_A/M",
                         RESET := "Pumps Data".R7_AG01.RESET,
                         "WAITING TIME" := "Pumps Data".R7_AG01.WT_SP,
                         OP_FBK_ERROR => "Valves Data".R7_VALVE_FAULT."AG01_FAIL_TO RUN",
                         "START/STOPCMD" => "DO_OUTPUT".R7_OUTPUTS."A/SSR_007_MOTOR",
                         STATUS => "Pumps Data".R7_AG01.STATUS);
   END_IF;
END_REGION

REGION Network 27: ***R8****
END_REGION

REGION Network 28: CP01
   RUNG wire#powerrail
      Contact( "AlwaysTRUE" )
      #PUMP_FB1_R8_CP01("AUTO START" := wire#w1, "PUMP SELECTION" := 1, TRIP := "A/SSR_008_CP01_TRIP_FB", SIM :=, "MANUAL SELECTION" := "Valves Data"."A/M".R8, SEMI :=, "MANUAL START" := "Pumps Data".R8_CP01.MCMD, "FEEDBACK RUN" := "A/SSR_008_CP01_RUN_FB", TRIPPED :=, REMOTE := "A/SSR_008_CP01_RL", RESET := "R8_DATA".R8.Reset, INTERLOCK :=, "WAITING TIME" := "Pumps Data".R8_CP01.WT_SP, OP_FBK_ERROR => "Valves Data".R8_VALVE_FAULT.CP01_FAIL_TO_RUN, CL_FBK_ERROR =>, AUTO_MODE =>, MANUAL_MODE =>, SEMI_AUTO_MODE =>, "START/STOPCMD" => "A/SSR_008_CP01_CMD", STATUS => "Pumps Data".R8_CP01.STATUS, FAULT =>)
   END_RUNG
   RUNG wire#powerrail
      Contact( "R8_DATA".R8.PUMP_CMD )
   END_RUNG wire#w1
   RUNG wire#powerrail
      Contact( "R8_DATA".R8.COOL_PUMP_CMD )
   END_RUNG wire#w1
   // the same network as SCL:
   IF "AlwaysTRUE" THEN
       #PUMP_FB1_R8_CP01("PUMP SELECTION" := 1,   // "PUMP_FB1"
                         TRIP := "A/SSR_008_CP01_TRIP_FB",
                         "AUTO START" := "R8_DATA".R8.PUMP_CMD OR "R8_DATA".R8.COOL_PUMP_CMD,
                         "MANUAL SELECTION" := "Valves Data"."A/M".R8,
                         "MANUAL START" := "Pumps Data".R8_CP01.MCMD,
                         "FEEDBACK RUN" := "A/SSR_008_CP01_RUN_FB",
                         REMOTE := "A/SSR_008_CP01_RL",
                         RESET := "R8_DATA".R8.Reset,
                         "WAITING TIME" := "Pumps Data".R8_CP01.WT_SP,
                         OP_FBK_ERROR => "Valves Data".R8_VALVE_FAULT.CP01_FAIL_TO_RUN,
                         "START/STOPCMD" => "A/SSR_008_CP01_CMD",
                         STATUS => "Pumps Data".R8_CP01.STATUS);
   END_IF;
END_REGION

REGION Network 29: AG01
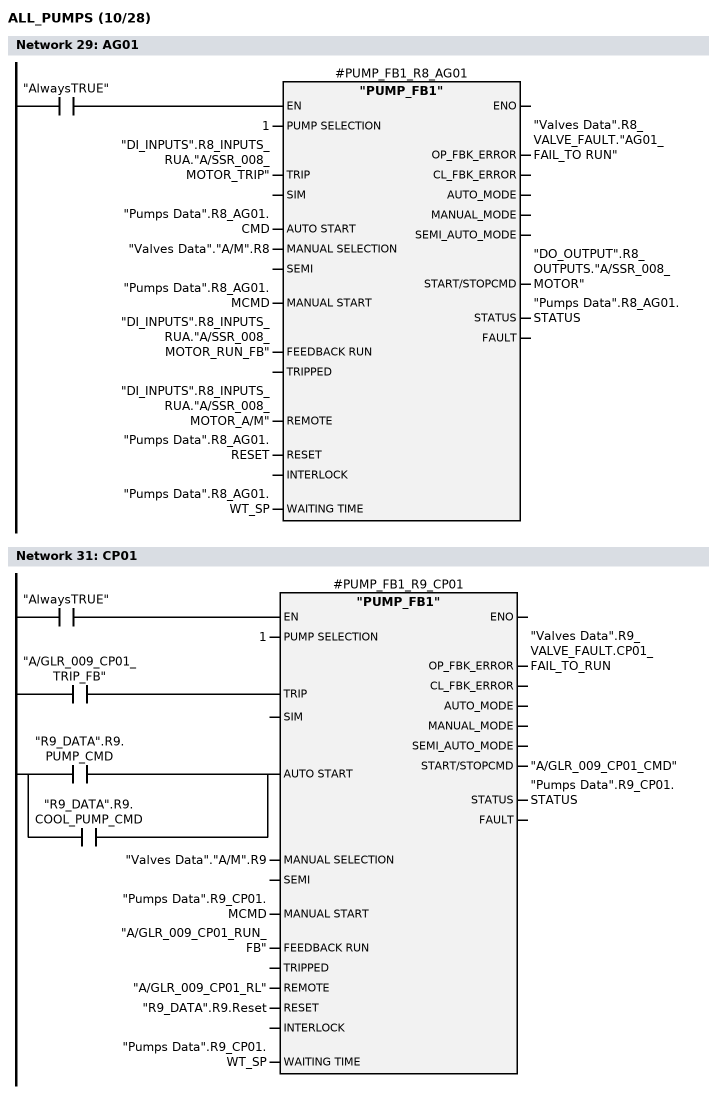
   RUNG wire#powerrail
      Contact( "AlwaysTRUE" )
      #PUMP_FB1_R8_AG01("PUMP SELECTION" := 1, TRIP := "DI_INPUTS".R8_INPUTS_RUA."A/SSR_008_MOTOR_TRIP", SIM :=, "AUTO START" := "Pumps Data".R8_AG01.CMD, "MANUAL SELECTION" := "Valves Data"."A/M".R8, SEMI :=, "MANUAL START" := "Pumps Data".R8_AG01.MCMD, "FEEDBACK RUN" := "DI_INPUTS".R8_INPUTS_RUA."A/SSR_008_MOTOR_RUN_FB", TRIPPED :=, REMOTE := "DI_INPUTS".R8_INPUTS_RUA."A/SSR_008_MOTOR_A/M", RESET := "Pumps Data".R8_AG01.RESET, INTERLOCK :=, "WAITING TIME" := "Pumps Data".R8_AG01.WT_SP, OP_FBK_ERROR => "Valves Data".R8_VALVE_FAULT."AG01_FAIL_TO RUN", CL_FBK_ERROR =>, AUTO_MODE =>, MANUAL_MODE =>, SEMI_AUTO_MODE =>, "START/STOPCMD" => "DO_OUTPUT".R8_OUTPUTS."A/SSR_008_MOTOR", STATUS => "Pumps Data".R8_AG01.STATUS, FAULT =>)
   END_RUNG
   // the same network as SCL:
   IF "AlwaysTRUE" THEN
       #PUMP_FB1_R8_AG01("PUMP SELECTION" := 1,   // "PUMP_FB1"
                         TRIP := "DI_INPUTS".R8_INPUTS_RUA."A/SSR_008_MOTOR_TRIP",
                         "AUTO START" := "Pumps Data".R8_AG01.CMD,
                         "MANUAL SELECTION" := "Valves Data"."A/M".R8,
                         "MANUAL START" := "Pumps Data".R8_AG01.MCMD,
                         "FEEDBACK RUN" := "DI_INPUTS".R8_INPUTS_RUA."A/SSR_008_MOTOR_RUN_FB",
                         REMOTE := "DI_INPUTS".R8_INPUTS_RUA."A/SSR_008_MOTOR_A/M",
                         RESET := "Pumps Data".R8_AG01.RESET,
                         "WAITING TIME" := "Pumps Data".R8_AG01.WT_SP,
                         OP_FBK_ERROR => "Valves Data".R8_VALVE_FAULT."AG01_FAIL_TO RUN",
                         "START/STOPCMD" => "DO_OUTPUT".R8_OUTPUTS."A/SSR_008_MOTOR",
                         STATUS => "Pumps Data".R8_AG01.STATUS);
   END_IF;
END_REGION

REGION Network 30: ***R9****
END_REGION

REGION Network 31: CP01
   RUNG wire#powerrail
      Contact( "AlwaysTRUE" )
      #PUMP_FB1_R9_CP01(TRIP := wire#w1, "AUTO START" := wire#w2, "PUMP SELECTION" := 1, SIM :=, "MANUAL SELECTION" := "Valves Data"."A/M".R9, SEMI :=, "MANUAL START" := "Pumps Data".R9_CP01.MCMD, "FEEDBACK RUN" := "A/GLR_009_CP01_RUN_FB", TRIPPED :=, REMOTE := "A/GLR_009_CP01_RL", RESET := "R9_DATA".R9.Reset, INTERLOCK :=, "WAITING TIME" := "Pumps Data".R9_CP01.WT_SP, OP_FBK_ERROR => "Valves Data".R9_VALVE_FAULT.CP01_FAIL_TO_RUN, CL_FBK_ERROR =>, AUTO_MODE =>, MANUAL_MODE =>, SEMI_AUTO_MODE =>, "START/STOPCMD" => "A/GLR_009_CP01_CMD", STATUS => "Pumps Data".R9_CP01.STATUS, FAULT =>)
   END_RUNG
   RUNG wire#powerrail
      Contact( "A/GLR_009_CP01_TRIP_FB" )
   END_RUNG wire#w1
   RUNG wire#powerrail
      Contact( "R9_DATA".R9.PUMP_CMD )
   END_RUNG wire#w2
   RUNG wire#powerrail
      Contact( "R9_DATA".R9.COOL_PUMP_CMD )
   END_RUNG wire#w2
   // the same network as SCL:
   IF "AlwaysTRUE" THEN
       #PUMP_FB1_R9_CP01("PUMP SELECTION" := 1,   // "PUMP_FB1"
                         TRIP := "A/GLR_009_CP01_TRIP_FB",
                         "AUTO START" := "R9_DATA".R9.PUMP_CMD OR "R9_DATA".R9.COOL_PUMP_CMD,
                         "MANUAL SELECTION" := "Valves Data"."A/M".R9,
                         "MANUAL START" := "Pumps Data".R9_CP01.MCMD,
                         "FEEDBACK RUN" := "A/GLR_009_CP01_RUN_FB",
                         REMOTE := "A/GLR_009_CP01_RL",
                         RESET := "R9_DATA".R9.Reset,
                         "WAITING TIME" := "Pumps Data".R9_CP01.WT_SP,
                         OP_FBK_ERROR => "Valves Data".R9_VALVE_FAULT.CP01_FAIL_TO_RUN,
                         "START/STOPCMD" => "A/GLR_009_CP01_CMD",
                         STATUS => "Pumps Data".R9_CP01.STATUS);
   END_IF;
END_REGION

REGION Network 32: AG01
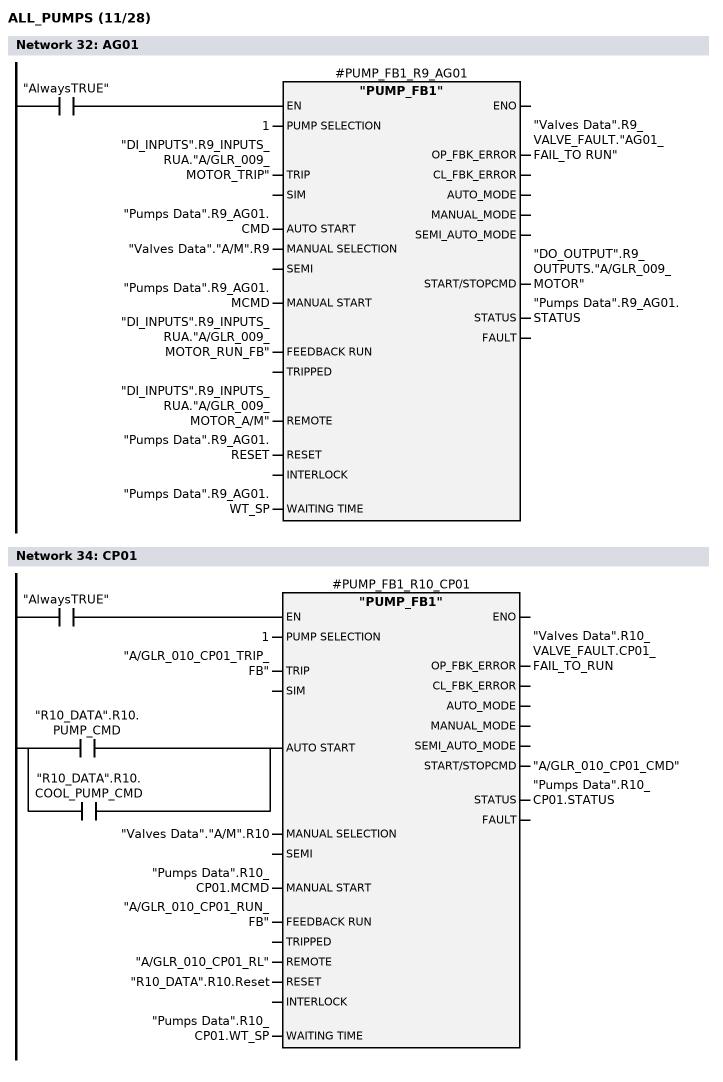
   RUNG wire#powerrail
      Contact( "AlwaysTRUE" )
      #PUMP_FB1_R9_AG01("PUMP SELECTION" := 1, TRIP := "DI_INPUTS".R9_INPUTS_RUA."A/GLR_009_MOTOR_TRIP", SIM :=, "AUTO START" := "Pumps Data".R9_AG01.CMD, "MANUAL SELECTION" := "Valves Data"."A/M".R9, SEMI :=, "MANUAL START" := "Pumps Data".R9_AG01.MCMD, "FEEDBACK RUN" := "DI_INPUTS".R9_INPUTS_RUA."A/GLR_009_MOTOR_RUN_FB", TRIPPED :=, REMOTE := "DI_INPUTS".R9_INPUTS_RUA."A/GLR_009_MOTOR_A/M", RESET := "Pumps Data".R9_AG01.RESET, INTERLOCK :=, "WAITING TIME" := "Pumps Data".R9_AG01.WT_SP, OP_FBK_ERROR => "Valves Data".R9_VALVE_FAULT."AG01_FAIL_TO RUN", CL_FBK_ERROR =>, AUTO_MODE =>, MANUAL_MODE =>, SEMI_AUTO_MODE =>, "START/STOPCMD" => "DO_OUTPUT".R9_OUTPUTS."A/GLR_009_MOTOR", STATUS => "Pumps Data".R9_AG01.STATUS, FAULT =>)
   END_RUNG
   // the same network as SCL:
   IF "AlwaysTRUE" THEN
       #PUMP_FB1_R9_AG01("PUMP SELECTION" := 1,   // "PUMP_FB1"
                         TRIP := "DI_INPUTS".R9_INPUTS_RUA."A/GLR_009_MOTOR_TRIP",
                         "AUTO START" := "Pumps Data".R9_AG01.CMD,
                         "MANUAL SELECTION" := "Valves Data"."A/M".R9,
                         "MANUAL START" := "Pumps Data".R9_AG01.MCMD,
                         "FEEDBACK RUN" := "DI_INPUTS".R9_INPUTS_RUA."A/GLR_009_MOTOR_RUN_FB",
                         REMOTE := "DI_INPUTS".R9_INPUTS_RUA."A/GLR_009_MOTOR_A/M",
                         RESET := "Pumps Data".R9_AG01.RESET,
                         "WAITING TIME" := "Pumps Data".R9_AG01.WT_SP,
                         OP_FBK_ERROR => "Valves Data".R9_VALVE_FAULT."AG01_FAIL_TO RUN",
                         "START/STOPCMD" => "DO_OUTPUT".R9_OUTPUTS."A/GLR_009_MOTOR",
                         STATUS => "Pumps Data".R9_AG01.STATUS);
   END_IF;
END_REGION

REGION Network 33: ***R10****
END_REGION

REGION Network 34: CP01
   RUNG wire#powerrail
      Contact( "AlwaysTRUE" )
      #PUMP_FB1_R10_CP01("AUTO START" := wire#w1, "PUMP SELECTION" := 1, TRIP := "A/GLR_010_CP01_TRIP_FB", SIM :=, "MANUAL SELECTION" := "Valves Data"."A/M".R10, SEMI :=, "MANUAL START" := "Pumps Data".R10_CP01.MCMD, "FEEDBACK RUN" := "A/GLR_010_CP01_RUN_FB", TRIPPED :=, REMOTE := "A/GLR_010_CP01_RL", RESET := "R10_DATA".R10.Reset, INTERLOCK :=, "WAITING TIME" := "Pumps Data".R10_CP01.WT_SP, OP_FBK_ERROR => "Valves Data".R10_VALVE_FAULT.CP01_FAIL_TO_RUN, CL_FBK_ERROR =>, AUTO_MODE =>, MANUAL_MODE =>, SEMI_AUTO_MODE =>, "START/STOPCMD" => "A/GLR_010_CP01_CMD", STATUS => "Pumps Data".R10_CP01.STATUS, FAULT =>)
   END_RUNG
   RUNG wire#powerrail
      Contact( "R10_DATA".R10.PUMP_CMD )
   END_RUNG wire#w1
   RUNG wire#powerrail
      Contact( "R10_DATA".R10.COOL_PUMP_CMD )
   END_RUNG wire#w1
   // the same network as SCL:
   IF "AlwaysTRUE" THEN
       #PUMP_FB1_R10_CP01("PUMP SELECTION" := 1,   // "PUMP_FB1"
                          TRIP := "A/GLR_010_CP01_TRIP_FB",
                          "AUTO START" := "R10_DATA".R10.PUMP_CMD OR "R10_DATA".R10.COOL_PUMP_CMD,
                          "MANUAL SELECTION" := "Valves Data"."A/M".R10,
                          "MANUAL START" := "Pumps Data".R10_CP01.MCMD,
                          "FEEDBACK RUN" := "A/GLR_010_CP01_RUN_FB",
                          REMOTE := "A/GLR_010_CP01_RL",
                          RESET := "R10_DATA".R10.Reset,
                          "WAITING TIME" := "Pumps Data".R10_CP01.WT_SP,
                          OP_FBK_ERROR => "Valves Data".R10_VALVE_FAULT.CP01_FAIL_TO_RUN,
                          "START/STOPCMD" => "A/GLR_010_CP01_CMD",
                          STATUS => "Pumps Data".R10_CP01.STATUS);
   END_IF;
END_REGION

REGION Network 35: AG01
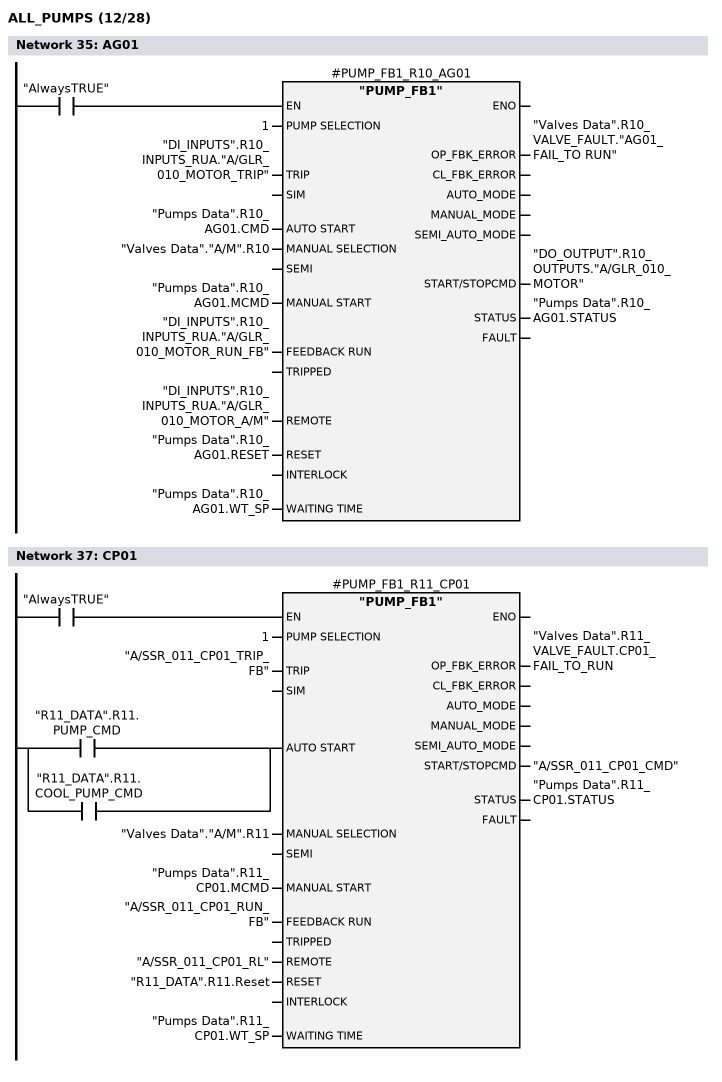
   RUNG wire#powerrail
      Contact( "AlwaysTRUE" )
      #PUMP_FB1_R10_AG01("PUMP SELECTION" := 1, TRIP := "DI_INPUTS".R10_INPUTS_RUA."A/GLR_010_MOTOR_TRIP", SIM :=, "AUTO START" := "Pumps Data".R10_AG01.CMD, "MANUAL SELECTION" := "Valves Data"."A/M".R10, SEMI :=, "MANUAL START" := "Pumps Data".R10_AG01.MCMD, "FEEDBACK RUN" := "DI_INPUTS".R10_INPUTS_RUA."A/GLR_010_MOTOR_RUN_FB", TRIPPED :=, REMOTE := "DI_INPUTS".R10_INPUTS_RUA."A/GLR_010_MOTOR_A/M", RESET := "Pumps Data".R10_AG01.RESET, INTERLOCK :=, "WAITING TIME" := "Pumps Data".R10_AG01.WT_SP, OP_FBK_ERROR => "Valves Data".R10_VALVE_FAULT."AG01_FAIL_TO RUN", CL_FBK_ERROR =>, AUTO_MODE =>, MANUAL_MODE =>, SEMI_AUTO_MODE =>, "START/STOPCMD" => "DO_OUTPUT".R10_OUTPUTS."A/GLR_010_MOTOR", STATUS => "Pumps Data".R10_AG01.STATUS, FAULT =>)
   END_RUNG
   // the same network as SCL:
   IF "AlwaysTRUE" THEN
       #PUMP_FB1_R10_AG01("PUMP SELECTION" := 1,   // "PUMP_FB1"
                          TRIP := "DI_INPUTS".R10_INPUTS_RUA."A/GLR_010_MOTOR_TRIP",
                          "AUTO START" := "Pumps Data".R10_AG01.CMD,
                          "MANUAL SELECTION" := "Valves Data"."A/M".R10,
                          "MANUAL START" := "Pumps Data".R10_AG01.MCMD,
                          "FEEDBACK RUN" := "DI_INPUTS".R10_INPUTS_RUA."A/GLR_010_MOTOR_RUN_FB",
                          REMOTE := "DI_INPUTS".R10_INPUTS_RUA."A/GLR_010_MOTOR_A/M",
                          RESET := "Pumps Data".R10_AG01.RESET,
                          "WAITING TIME" := "Pumps Data".R10_AG01.WT_SP,
                          OP_FBK_ERROR => "Valves Data".R10_VALVE_FAULT."AG01_FAIL_TO RUN",
                          "START/STOPCMD" => "DO_OUTPUT".R10_OUTPUTS."A/GLR_010_MOTOR",
                          STATUS => "Pumps Data".R10_AG01.STATUS);
   END_IF;
END_REGION

REGION Network 36: ***R11****
END_REGION

REGION Network 37: CP01
   RUNG wire#powerrail
      Contact( "AlwaysTRUE" )
      #PUMP_FB1_R11_CP01("AUTO START" := wire#w1, "PUMP SELECTION" := 1, TRIP := "A/SSR_011_CP01_TRIP_FB", SIM :=, "MANUAL SELECTION" := "Valves Data"."A/M".R11, SEMI :=, "MANUAL START" := "Pumps Data".R11_CP01.MCMD, "FEEDBACK RUN" := "A/SSR_011_CP01_RUN_FB", TRIPPED :=, REMOTE := "A/SSR_011_CP01_RL", RESET := "R11_DATA".R11.Reset, INTERLOCK :=, "WAITING TIME" := "Pumps Data".R11_CP01.WT_SP, OP_FBK_ERROR => "Valves Data".R11_VALVE_FAULT.CP01_FAIL_TO_RUN, CL_FBK_ERROR =>, AUTO_MODE =>, MANUAL_MODE =>, SEMI_AUTO_MODE =>, "START/STOPCMD" => "A/SSR_011_CP01_CMD", STATUS => "Pumps Data".R11_CP01.STATUS, FAULT =>)
   END_RUNG
   RUNG wire#powerrail
      Contact( "R11_DATA".R11.PUMP_CMD )
   END_RUNG wire#w1
   RUNG wire#powerrail
      Contact( "R11_DATA".R11.COOL_PUMP_CMD )
   END_RUNG wire#w1
   // the same network as SCL:
   IF "AlwaysTRUE" THEN
       #PUMP_FB1_R11_CP01("PUMP SELECTION" := 1,   // "PUMP_FB1"
                          TRIP := "A/SSR_011_CP01_TRIP_FB",
                          "AUTO START" := "R11_DATA".R11.PUMP_CMD OR "R11_DATA".R11.COOL_PUMP_CMD,
                          "MANUAL SELECTION" := "Valves Data"."A/M".R11,
                          "MANUAL START" := "Pumps Data".R11_CP01.MCMD,
                          "FEEDBACK RUN" := "A/SSR_011_CP01_RUN_FB",
                          REMOTE := "A/SSR_011_CP01_RL",
                          RESET := "R11_DATA".R11.Reset,
                          "WAITING TIME" := "Pumps Data".R11_CP01.WT_SP,
                          OP_FBK_ERROR => "Valves Data".R11_VALVE_FAULT.CP01_FAIL_TO_RUN,
                          "START/STOPCMD" => "A/SSR_011_CP01_CMD",
                          STATUS => "Pumps Data".R11_CP01.STATUS);
   END_IF;
END_REGION

REGION Network 38: AG01
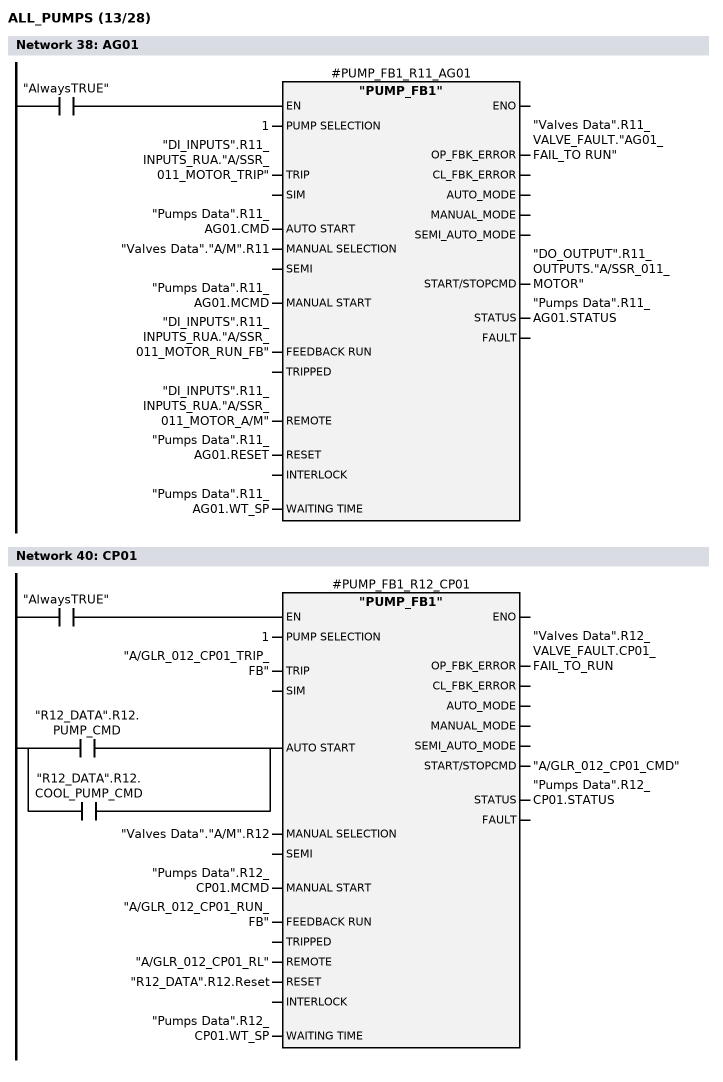
   RUNG wire#powerrail
      Contact( "AlwaysTRUE" )
      #PUMP_FB1_R11_AG01("PUMP SELECTION" := 1, TRIP := "DI_INPUTS".R11_INPUTS_RUA."A/SSR_011_MOTOR_TRIP", SIM :=, "AUTO START" := "Pumps Data".R11_AG01.CMD, "MANUAL SELECTION" := "Valves Data"."A/M".R11, SEMI :=, "MANUAL START" := "Pumps Data".R11_AG01.MCMD, "FEEDBACK RUN" := "DI_INPUTS".R11_INPUTS_RUA."A/SSR_011_MOTOR_RUN_FB", TRIPPED :=, REMOTE := "DI_INPUTS".R11_INPUTS_RUA."A/SSR_011_MOTOR_A/M", RESET := "Pumps Data".R11_AG01.RESET, INTERLOCK :=, "WAITING TIME" := "Pumps Data".R11_AG01.WT_SP, OP_FBK_ERROR => "Valves Data".R11_VALVE_FAULT."AG01_FAIL_TO RUN", CL_FBK_ERROR =>, AUTO_MODE =>, MANUAL_MODE =>, SEMI_AUTO_MODE =>, "START/STOPCMD" => "DO_OUTPUT".R11_OUTPUTS."A/SSR_011_MOTOR", STATUS => "Pumps Data".R11_AG01.STATUS, FAULT =>)
   END_RUNG
   // the same network as SCL:
   IF "AlwaysTRUE" THEN
       #PUMP_FB1_R11_AG01("PUMP SELECTION" := 1,   // "PUMP_FB1"
                          TRIP := "DI_INPUTS".R11_INPUTS_RUA."A/SSR_011_MOTOR_TRIP",
                          "AUTO START" := "Pumps Data".R11_AG01.CMD,
                          "MANUAL SELECTION" := "Valves Data"."A/M".R11,
                          "MANUAL START" := "Pumps Data".R11_AG01.MCMD,
                          "FEEDBACK RUN" := "DI_INPUTS".R11_INPUTS_RUA."A/SSR_011_MOTOR_RUN_FB",
                          REMOTE := "DI_INPUTS".R11_INPUTS_RUA."A/SSR_011_MOTOR_A/M",
                          RESET := "Pumps Data".R11_AG01.RESET,
                          "WAITING TIME" := "Pumps Data".R11_AG01.WT_SP,
                          OP_FBK_ERROR => "Valves Data".R11_VALVE_FAULT."AG01_FAIL_TO RUN",
                          "START/STOPCMD" => "DO_OUTPUT".R11_OUTPUTS."A/SSR_011_MOTOR",
                          STATUS => "Pumps Data".R11_AG01.STATUS);
   END_IF;
END_REGION

REGION Network 39: ***R12****
END_REGION

REGION Network 40: CP01
   RUNG wire#powerrail
      Contact( "AlwaysTRUE" )
      #PUMP_FB1_R12_CP01("AUTO START" := wire#w1, "PUMP SELECTION" := 1, TRIP := "A/GLR_012_CP01_TRIP_FB", SIM :=, "MANUAL SELECTION" := "Valves Data"."A/M".R12, SEMI :=, "MANUAL START" := "Pumps Data".R12_CP01.MCMD, "FEEDBACK RUN" := "A/GLR_012_CP01_RUN_FB", TRIPPED :=, REMOTE := "A/GLR_012_CP01_RL", RESET := "R12_DATA".R12.Reset, INTERLOCK :=, "WAITING TIME" := "Pumps Data".R12_CP01.WT_SP, OP_FBK_ERROR => "Valves Data".R12_VALVE_FAULT.CP01_FAIL_TO_RUN, CL_FBK_ERROR =>, AUTO_MODE =>, MANUAL_MODE =>, SEMI_AUTO_MODE =>, "START/STOPCMD" => "A/GLR_012_CP01_CMD", STATUS => "Pumps Data".R12_CP01.STATUS, FAULT =>)
   END_RUNG
   RUNG wire#powerrail
      Contact( "R12_DATA".R12.PUMP_CMD )
   END_RUNG wire#w1
   RUNG wire#powerrail
      Contact( "R12_DATA".R12.COOL_PUMP_CMD )
   END_RUNG wire#w1
   // the same network as SCL:
   IF "AlwaysTRUE" THEN
       #PUMP_FB1_R12_CP01("PUMP SELECTION" := 1,   // "PUMP_FB1"
                          TRIP := "A/GLR_012_CP01_TRIP_FB",
                          "AUTO START" := "R12_DATA".R12.PUMP_CMD OR "R12_DATA".R12.COOL_PUMP_CMD,
                          "MANUAL SELECTION" := "Valves Data"."A/M".R12,
                          "MANUAL START" := "Pumps Data".R12_CP01.MCMD,
                          "FEEDBACK RUN" := "A/GLR_012_CP01_RUN_FB",
                          REMOTE := "A/GLR_012_CP01_RL",
                          RESET := "R12_DATA".R12.Reset,
                          "WAITING TIME" := "Pumps Data".R12_CP01.WT_SP,
                          OP_FBK_ERROR => "Valves Data".R12_VALVE_FAULT.CP01_FAIL_TO_RUN,
                          "START/STOPCMD" => "A/GLR_012_CP01_CMD",
                          STATUS => "Pumps Data".R12_CP01.STATUS);
   END_IF;
END_REGION

REGION Network 41: AG01
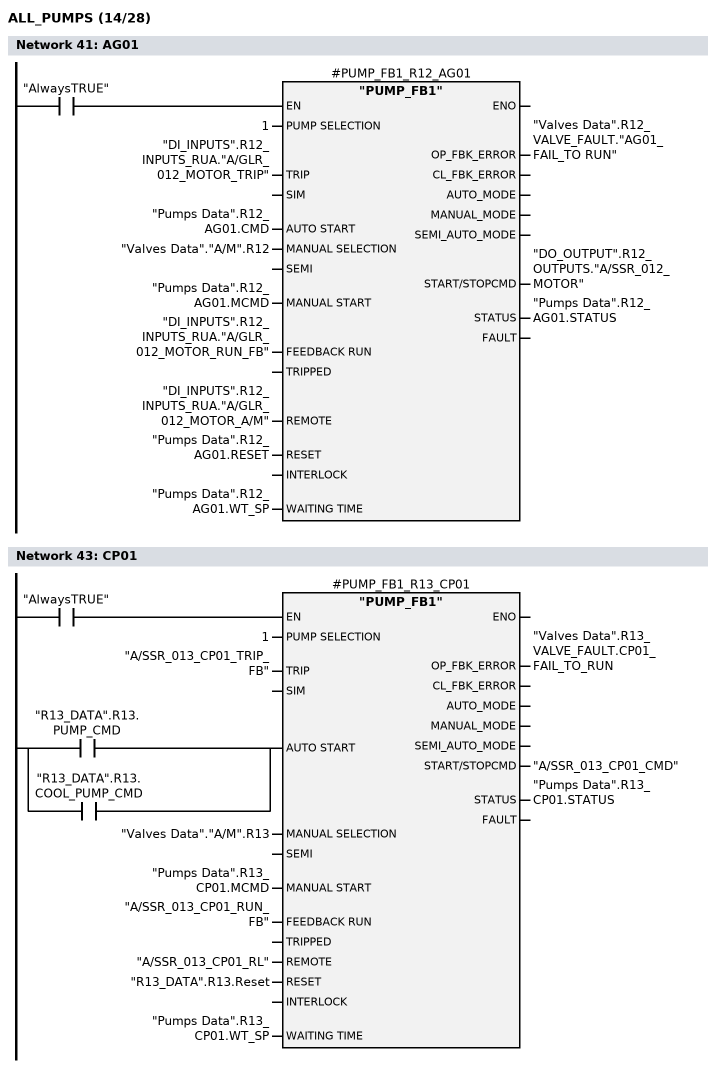
   RUNG wire#powerrail
      Contact( "AlwaysTRUE" )
      #PUMP_FB1_R12_AG01("PUMP SELECTION" := 1, TRIP := "DI_INPUTS".R12_INPUTS_RUA."A/GLR_012_MOTOR_TRIP", SIM :=, "AUTO START" := "Pumps Data".R12_AG01.CMD, "MANUAL SELECTION" := "Valves Data"."A/M".R12, SEMI :=, "MANUAL START" := "Pumps Data".R12_AG01.MCMD, "FEEDBACK RUN" := "DI_INPUTS".R12_INPUTS_RUA."A/GLR_012_MOTOR_RUN_FB", TRIPPED :=, REMOTE := "DI_INPUTS".R12_INPUTS_RUA."A/GLR_012_MOTOR_A/M", RESET := "Pumps Data".R12_AG01.RESET, INTERLOCK :=, "WAITING TIME" := "Pumps Data".R12_AG01.WT_SP, OP_FBK_ERROR => "Valves Data".R12_VALVE_FAULT."AG01_FAIL_TO RUN", CL_FBK_ERROR =>, AUTO_MODE =>, MANUAL_MODE =>, SEMI_AUTO_MODE =>, "START/STOPCMD" => "DO_OUTPUT".R12_OUTPUTS."A/SSR_012_MOTOR", STATUS => "Pumps Data".R12_AG01.STATUS, FAULT =>)
   END_RUNG
   // the same network as SCL:
   IF "AlwaysTRUE" THEN
       #PUMP_FB1_R12_AG01("PUMP SELECTION" := 1,   // "PUMP_FB1"
                          TRIP := "DI_INPUTS".R12_INPUTS_RUA."A/GLR_012_MOTOR_TRIP",
                          "AUTO START" := "Pumps Data".R12_AG01.CMD,
                          "MANUAL SELECTION" := "Valves Data"."A/M".R12,
                          "MANUAL START" := "Pumps Data".R12_AG01.MCMD,
                          "FEEDBACK RUN" := "DI_INPUTS".R12_INPUTS_RUA."A/GLR_012_MOTOR_RUN_FB",
                          REMOTE := "DI_INPUTS".R12_INPUTS_RUA."A/GLR_012_MOTOR_A/M",
                          RESET := "Pumps Data".R12_AG01.RESET,
                          "WAITING TIME" := "Pumps Data".R12_AG01.WT_SP,
                          OP_FBK_ERROR => "Valves Data".R12_VALVE_FAULT."AG01_FAIL_TO RUN",
                          "START/STOPCMD" => "DO_OUTPUT".R12_OUTPUTS."A/SSR_012_MOTOR",
                          STATUS => "Pumps Data".R12_AG01.STATUS);
   END_IF;
END_REGION

REGION Network 42: ***R13****
END_REGION

REGION Network 43: CP01
   RUNG wire#powerrail
      Contact( "AlwaysTRUE" )
      #PUMP_FB1_R13_CP01("AUTO START" := wire#w1, "PUMP SELECTION" := 1, TRIP := "A/SSR_013_CP01_TRIP_FB", SIM :=, "MANUAL SELECTION" := "Valves Data"."A/M".R13, SEMI :=, "MANUAL START" := "Pumps Data".R13_CP01.MCMD, "FEEDBACK RUN" := "A/SSR_013_CP01_RUN_FB", TRIPPED :=, REMOTE := "A/SSR_013_CP01_RL", RESET := "R13_DATA".R13.Reset, INTERLOCK :=, "WAITING TIME" := "Pumps Data".R13_CP01.WT_SP, OP_FBK_ERROR => "Valves Data".R13_VALVE_FAULT.CP01_FAIL_TO_RUN, CL_FBK_ERROR =>, AUTO_MODE =>, MANUAL_MODE =>, SEMI_AUTO_MODE =>, "START/STOPCMD" => "A/SSR_013_CP01_CMD", STATUS => "Pumps Data".R13_CP01.STATUS, FAULT =>)
   END_RUNG
   RUNG wire#powerrail
      Contact( "R13_DATA".R13.PUMP_CMD )
   END_RUNG wire#w1
   RUNG wire#powerrail
      Contact( "R13_DATA".R13.COOL_PUMP_CMD )
   END_RUNG wire#w1
   // the same network as SCL:
   IF "AlwaysTRUE" THEN
       #PUMP_FB1_R13_CP01("PUMP SELECTION" := 1,   // "PUMP_FB1"
                          TRIP := "A/SSR_013_CP01_TRIP_FB",
                          "AUTO START" := "R13_DATA".R13.PUMP_CMD OR "R13_DATA".R13.COOL_PUMP_CMD,
                          "MANUAL SELECTION" := "Valves Data"."A/M".R13,
                          "MANUAL START" := "Pumps Data".R13_CP01.MCMD,
                          "FEEDBACK RUN" := "A/SSR_013_CP01_RUN_FB",
                          REMOTE := "A/SSR_013_CP01_RL",
                          RESET := "R13_DATA".R13.Reset,
                          "WAITING TIME" := "Pumps Data".R13_CP01.WT_SP,
                          OP_FBK_ERROR => "Valves Data".R13_VALVE_FAULT.CP01_FAIL_TO_RUN,
                          "START/STOPCMD" => "A/SSR_013_CP01_CMD",
                          STATUS => "Pumps Data".R13_CP01.STATUS);
   END_IF;
END_REGION

REGION Network 44: AG01
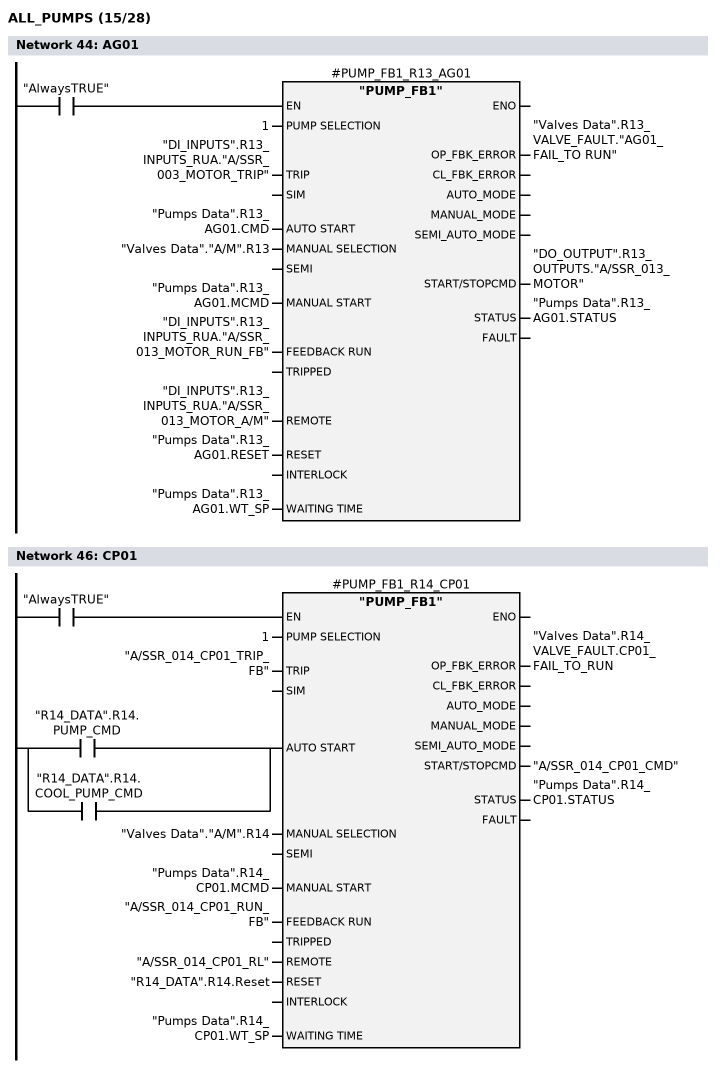
   RUNG wire#powerrail
      Contact( "AlwaysTRUE" )
      #PUMP_FB1_R13_AG01("PUMP SELECTION" := 1, TRIP := "DI_INPUTS".R13_INPUTS_RUA."A/SSR_003_MOTOR_TRIP", SIM :=, "AUTO START" := "Pumps Data".R13_AG01.CMD, "MANUAL SELECTION" := "Valves Data"."A/M".R13, SEMI :=, "MANUAL START" := "Pumps Data".R13_AG01.MCMD, "FEEDBACK RUN" := "DI_INPUTS".R13_INPUTS_RUA."A/SSR_013_MOTOR_RUN_FB", TRIPPED :=, REMOTE := "DI_INPUTS".R13_INPUTS_RUA."A/SSR_013_MOTOR_A/M", RESET := "Pumps Data".R13_AG01.RESET, INTERLOCK :=, "WAITING TIME" := "Pumps Data".R13_AG01.WT_SP, OP_FBK_ERROR => "Valves Data".R13_VALVE_FAULT."AG01_FAIL_TO RUN", CL_FBK_ERROR =>, AUTO_MODE =>, MANUAL_MODE =>, SEMI_AUTO_MODE =>, "START/STOPCMD" => "DO_OUTPUT".R13_OUTPUTS."A/SSR_013_MOTOR", STATUS => "Pumps Data".R13_AG01.STATUS, FAULT =>)
   END_RUNG
   // the same network as SCL:
   IF "AlwaysTRUE" THEN
       #PUMP_FB1_R13_AG01("PUMP SELECTION" := 1,   // "PUMP_FB1"
                          TRIP := "DI_INPUTS".R13_INPUTS_RUA."A/SSR_003_MOTOR_TRIP",
                          "AUTO START" := "Pumps Data".R13_AG01.CMD,
                          "MANUAL SELECTION" := "Valves Data"."A/M".R13,
                          "MANUAL START" := "Pumps Data".R13_AG01.MCMD,
                          "FEEDBACK RUN" := "DI_INPUTS".R13_INPUTS_RUA."A/SSR_013_MOTOR_RUN_FB",
                          REMOTE := "DI_INPUTS".R13_INPUTS_RUA."A/SSR_013_MOTOR_A/M",
                          RESET := "Pumps Data".R13_AG01.RESET,
                          "WAITING TIME" := "Pumps Data".R13_AG01.WT_SP,
                          OP_FBK_ERROR => "Valves Data".R13_VALVE_FAULT."AG01_FAIL_TO RUN",
                          "START/STOPCMD" => "DO_OUTPUT".R13_OUTPUTS."A/SSR_013_MOTOR",
                          STATUS => "Pumps Data".R13_AG01.STATUS);
   END_IF;
END_REGION

REGION Network 45: ***R14****
END_REGION

REGION Network 46: CP01
   RUNG wire#powerrail
      Contact( "AlwaysTRUE" )
      #PUMP_FB1_R14_CP01("AUTO START" := wire#w1, "PUMP SELECTION" := 1, TRIP := "A/SSR_014_CP01_TRIP_FB", SIM :=, "MANUAL SELECTION" := "Valves Data"."A/M".R14, SEMI :=, "MANUAL START" := "Pumps Data".R14_CP01.MCMD, "FEEDBACK RUN" := "A/SSR_014_CP01_RUN_FB", TRIPPED :=, REMOTE := "A/SSR_014_CP01_RL", RESET := "R14_DATA".R14.Reset, INTERLOCK :=, "WAITING TIME" := "Pumps Data".R14_CP01.WT_SP, OP_FBK_ERROR => "Valves Data".R14_VALVE_FAULT.CP01_FAIL_TO_RUN, CL_FBK_ERROR =>, AUTO_MODE =>, MANUAL_MODE =>, SEMI_AUTO_MODE =>, "START/STOPCMD" => "A/SSR_014_CP01_CMD", STATUS => "Pumps Data".R14_CP01.STATUS, FAULT =>)
   END_RUNG
   RUNG wire#powerrail
      Contact( "R14_DATA".R14.PUMP_CMD )
   END_RUNG wire#w1
   RUNG wire#powerrail
      Contact( "R14_DATA".R14.COOL_PUMP_CMD )
   END_RUNG wire#w1
   // the same network as SCL:
   IF "AlwaysTRUE" THEN
       #PUMP_FB1_R14_CP01("PUMP SELECTION" := 1,   // "PUMP_FB1"
                          TRIP := "A/SSR_014_CP01_TRIP_FB",
                          "AUTO START" := "R14_DATA".R14.PUMP_CMD OR "R14_DATA".R14.COOL_PUMP_CMD,
                          "MANUAL SELECTION" := "Valves Data"."A/M".R14,
                          "MANUAL START" := "Pumps Data".R14_CP01.MCMD,
                          "FEEDBACK RUN" := "A/SSR_014_CP01_RUN_FB",
                          REMOTE := "A/SSR_014_CP01_RL",
                          RESET := "R14_DATA".R14.Reset,
                          "WAITING TIME" := "Pumps Data".R14_CP01.WT_SP,
                          OP_FBK_ERROR => "Valves Data".R14_VALVE_FAULT.CP01_FAIL_TO_RUN,
                          "START/STOPCMD" => "A/SSR_014_CP01_CMD",
                          STATUS => "Pumps Data".R14_CP01.STATUS);
   END_IF;
END_REGION

REGION Network 47: AG01
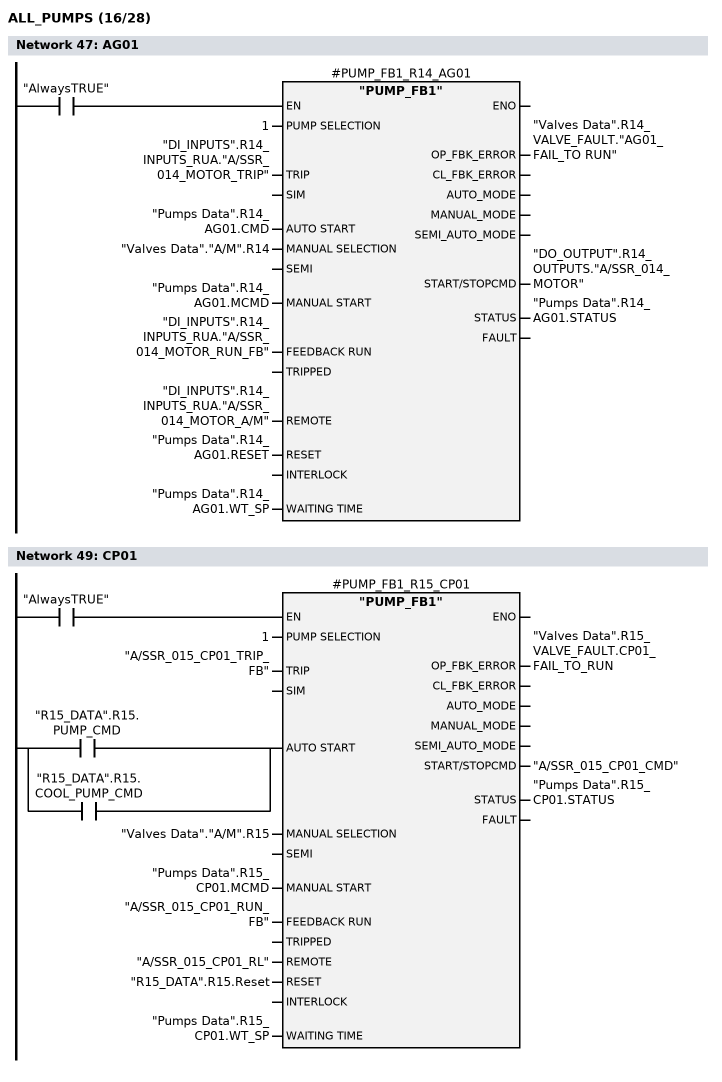
   RUNG wire#powerrail
      Contact( "AlwaysTRUE" )
      #PUMP_FB1_R14_AG01("PUMP SELECTION" := 1, TRIP := "DI_INPUTS".R14_INPUTS_RUA."A/SSR_014_MOTOR_TRIP", SIM :=, "AUTO START" := "Pumps Data".R14_AG01.CMD, "MANUAL SELECTION" := "Valves Data"."A/M".R14, SEMI :=, "MANUAL START" := "Pumps Data".R14_AG01.MCMD, "FEEDBACK RUN" := "DI_INPUTS".R14_INPUTS_RUA."A/SSR_014_MOTOR_RUN_FB", TRIPPED :=, REMOTE := "DI_INPUTS".R14_INPUTS_RUA."A/SSR_014_MOTOR_A/M", RESET := "Pumps Data".R14_AG01.RESET, INTERLOCK :=, "WAITING TIME" := "Pumps Data".R14_AG01.WT_SP, OP_FBK_ERROR => "Valves Data".R14_VALVE_FAULT."AG01_FAIL_TO RUN", CL_FBK_ERROR =>, AUTO_MODE =>, MANUAL_MODE =>, SEMI_AUTO_MODE =>, "START/STOPCMD" => "DO_OUTPUT".R14_OUTPUTS."A/SSR_014_MOTOR", STATUS => "Pumps Data".R14_AG01.STATUS, FAULT =>)
   END_RUNG
   // the same network as SCL:
   IF "AlwaysTRUE" THEN
       #PUMP_FB1_R14_AG01("PUMP SELECTION" := 1,   // "PUMP_FB1"
                          TRIP := "DI_INPUTS".R14_INPUTS_RUA."A/SSR_014_MOTOR_TRIP",
                          "AUTO START" := "Pumps Data".R14_AG01.CMD,
                          "MANUAL SELECTION" := "Valves Data"."A/M".R14,
                          "MANUAL START" := "Pumps Data".R14_AG01.MCMD,
                          "FEEDBACK RUN" := "DI_INPUTS".R14_INPUTS_RUA."A/SSR_014_MOTOR_RUN_FB",
                          REMOTE := "DI_INPUTS".R14_INPUTS_RUA."A/SSR_014_MOTOR_A/M",
                          RESET := "Pumps Data".R14_AG01.RESET,
                          "WAITING TIME" := "Pumps Data".R14_AG01.WT_SP,
                          OP_FBK_ERROR => "Valves Data".R14_VALVE_FAULT."AG01_FAIL_TO RUN",
                          "START/STOPCMD" => "DO_OUTPUT".R14_OUTPUTS."A/SSR_014_MOTOR",
                          STATUS => "Pumps Data".R14_AG01.STATUS);
   END_IF;
END_REGION

REGION Network 48: ***R15****
END_REGION

REGION Network 49: CP01
   RUNG wire#powerrail
      Contact( "AlwaysTRUE" )
      #PUMP_FB1_R15_CP01("AUTO START" := wire#w1, "PUMP SELECTION" := 1, TRIP := "A/SSR_015_CP01_TRIP_FB", SIM :=, "MANUAL SELECTION" := "Valves Data"."A/M".R15, SEMI :=, "MANUAL START" := "Pumps Data".R15_CP01.MCMD, "FEEDBACK RUN" := "A/SSR_015_CP01_RUN_FB", TRIPPED :=, REMOTE := "A/SSR_015_CP01_RL", RESET := "R15_DATA".R15.Reset, INTERLOCK :=, "WAITING TIME" := "Pumps Data".R15_CP01.WT_SP, OP_FBK_ERROR => "Valves Data".R15_VALVE_FAULT.CP01_FAIL_TO_RUN, CL_FBK_ERROR =>, AUTO_MODE =>, MANUAL_MODE =>, SEMI_AUTO_MODE =>, "START/STOPCMD" => "A/SSR_015_CP01_CMD", STATUS => "Pumps Data".R15_CP01.STATUS, FAULT =>)
   END_RUNG
   RUNG wire#powerrail
      Contact( "R15_DATA".R15.PUMP_CMD )
   END_RUNG wire#w1
   RUNG wire#powerrail
      Contact( "R15_DATA".R15.COOL_PUMP_CMD )
   END_RUNG wire#w1
   // the same network as SCL:
   IF "AlwaysTRUE" THEN
       #PUMP_FB1_R15_CP01("PUMP SELECTION" := 1,   // "PUMP_FB1"
                          TRIP := "A/SSR_015_CP01_TRIP_FB",
                          "AUTO START" := "R15_DATA".R15.PUMP_CMD OR "R15_DATA".R15.COOL_PUMP_CMD,
                          "MANUAL SELECTION" := "Valves Data"."A/M".R15,
                          "MANUAL START" := "Pumps Data".R15_CP01.MCMD,
                          "FEEDBACK RUN" := "A/SSR_015_CP01_RUN_FB",
                          REMOTE := "A/SSR_015_CP01_RL",
                          RESET := "R15_DATA".R15.Reset,
                          "WAITING TIME" := "Pumps Data".R15_CP01.WT_SP,
                          OP_FBK_ERROR => "Valves Data".R15_VALVE_FAULT.CP01_FAIL_TO_RUN,
                          "START/STOPCMD" => "A/SSR_015_CP01_CMD",
                          STATUS => "Pumps Data".R15_CP01.STATUS);
   END_IF;
END_REGION

REGION Network 50: AG01
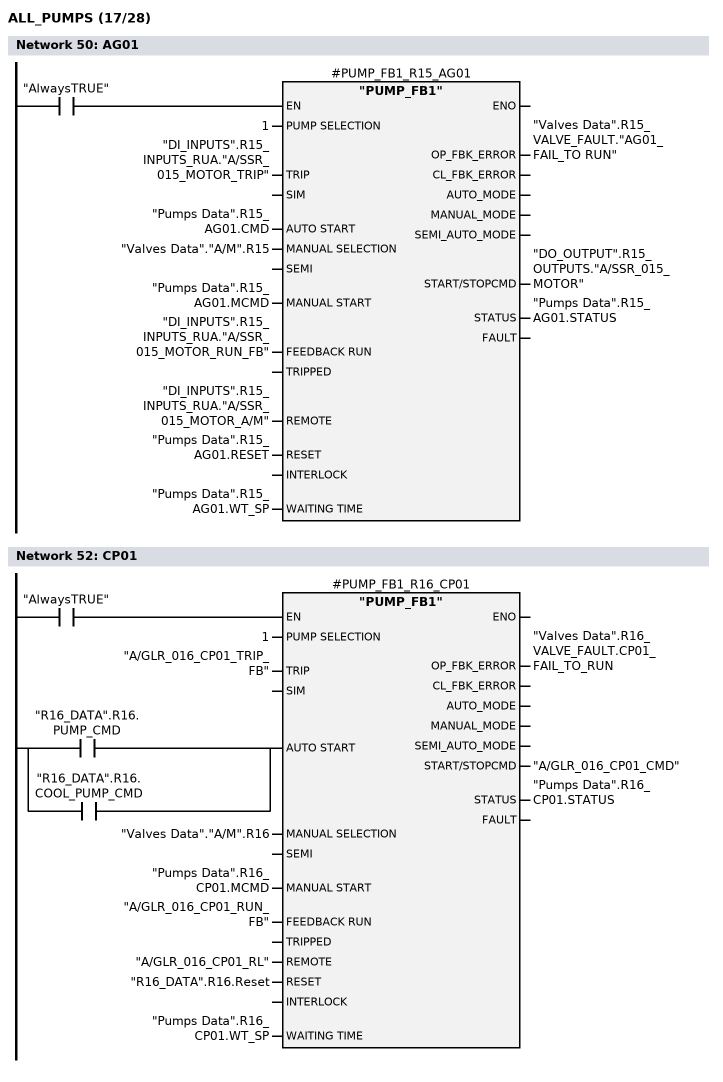
   RUNG wire#powerrail
      Contact( "AlwaysTRUE" )
      #PUMP_FB1_R15_AG01("PUMP SELECTION" := 1, TRIP := "DI_INPUTS".R15_INPUTS_RUA."A/SSR_015_MOTOR_TRIP", SIM :=, "AUTO START" := "Pumps Data".R15_AG01.CMD, "MANUAL SELECTION" := "Valves Data"."A/M".R15, SEMI :=, "MANUAL START" := "Pumps Data".R15_AG01.MCMD, "FEEDBACK RUN" := "DI_INPUTS".R15_INPUTS_RUA."A/SSR_015_MOTOR_RUN_FB", TRIPPED :=, REMOTE := "DI_INPUTS".R15_INPUTS_RUA."A/SSR_015_MOTOR_A/M", RESET := "Pumps Data".R15_AG01.RESET, INTERLOCK :=, "WAITING TIME" := "Pumps Data".R15_AG01.WT_SP, OP_FBK_ERROR => "Valves Data".R15_VALVE_FAULT."AG01_FAIL_TO RUN", CL_FBK_ERROR =>, AUTO_MODE =>, MANUAL_MODE =>, SEMI_AUTO_MODE =>, "START/STOPCMD" => "DO_OUTPUT".R15_OUTPUTS."A/SSR_015_MOTOR", STATUS => "Pumps Data".R15_AG01.STATUS, FAULT =>)
   END_RUNG
   // the same network as SCL:
   IF "AlwaysTRUE" THEN
       #PUMP_FB1_R15_AG01("PUMP SELECTION" := 1,   // "PUMP_FB1"
                          TRIP := "DI_INPUTS".R15_INPUTS_RUA."A/SSR_015_MOTOR_TRIP",
                          "AUTO START" := "Pumps Data".R15_AG01.CMD,
                          "MANUAL SELECTION" := "Valves Data"."A/M".R15,
                          "MANUAL START" := "Pumps Data".R15_AG01.MCMD,
                          "FEEDBACK RUN" := "DI_INPUTS".R15_INPUTS_RUA."A/SSR_015_MOTOR_RUN_FB",
                          REMOTE := "DI_INPUTS".R15_INPUTS_RUA."A/SSR_015_MOTOR_A/M",
                          RESET := "Pumps Data".R15_AG01.RESET,
                          "WAITING TIME" := "Pumps Data".R15_AG01.WT_SP,
                          OP_FBK_ERROR => "Valves Data".R15_VALVE_FAULT."AG01_FAIL_TO RUN",
                          "START/STOPCMD" => "DO_OUTPUT".R15_OUTPUTS."A/SSR_015_MOTOR",
                          STATUS => "Pumps Data".R15_AG01.STATUS);
   END_IF;
END_REGION

REGION Network 51: ***R16****
END_REGION

REGION Network 52: CP01
   RUNG wire#powerrail
      Contact( "AlwaysTRUE" )
      #PUMP_FB1_R16_CP01("AUTO START" := wire#w1, "PUMP SELECTION" := 1, TRIP := "A/GLR_016_CP01_TRIP_FB", SIM :=, "MANUAL SELECTION" := "Valves Data"."A/M".R16, SEMI :=, "MANUAL START" := "Pumps Data".R16_CP01.MCMD, "FEEDBACK RUN" := "A/GLR_016_CP01_RUN_FB", TRIPPED :=, REMOTE := "A/GLR_016_CP01_RL", RESET := "R16_DATA".R16.Reset, INTERLOCK :=, "WAITING TIME" := "Pumps Data".R16_CP01.WT_SP, OP_FBK_ERROR => "Valves Data".R16_VALVE_FAULT.CP01_FAIL_TO_RUN, CL_FBK_ERROR =>, AUTO_MODE =>, MANUAL_MODE =>, SEMI_AUTO_MODE =>, "START/STOPCMD" => "A/GLR_016_CP01_CMD", STATUS => "Pumps Data".R16_CP01.STATUS, FAULT =>)
   END_RUNG
   RUNG wire#powerrail
      Contact( "R16_DATA".R16.PUMP_CMD )
   END_RUNG wire#w1
   RUNG wire#powerrail
      Contact( "R16_DATA".R16.COOL_PUMP_CMD )
   END_RUNG wire#w1
   // the same network as SCL:
   IF "AlwaysTRUE" THEN
       #PUMP_FB1_R16_CP01("PUMP SELECTION" := 1,   // "PUMP_FB1"
                          TRIP := "A/GLR_016_CP01_TRIP_FB",
                          "AUTO START" := "R16_DATA".R16.PUMP_CMD OR "R16_DATA".R16.COOL_PUMP_CMD,
                          "MANUAL SELECTION" := "Valves Data"."A/M".R16,
                          "MANUAL START" := "Pumps Data".R16_CP01.MCMD,
                          "FEEDBACK RUN" := "A/GLR_016_CP01_RUN_FB",
                          REMOTE := "A/GLR_016_CP01_RL",
                          RESET := "R16_DATA".R16.Reset,
                          "WAITING TIME" := "Pumps Data".R16_CP01.WT_SP,
                          OP_FBK_ERROR => "Valves Data".R16_VALVE_FAULT.CP01_FAIL_TO_RUN,
                          "START/STOPCMD" => "A/GLR_016_CP01_CMD",
                          STATUS => "Pumps Data".R16_CP01.STATUS);
   END_IF;
END_REGION

REGION Network 53: AG01
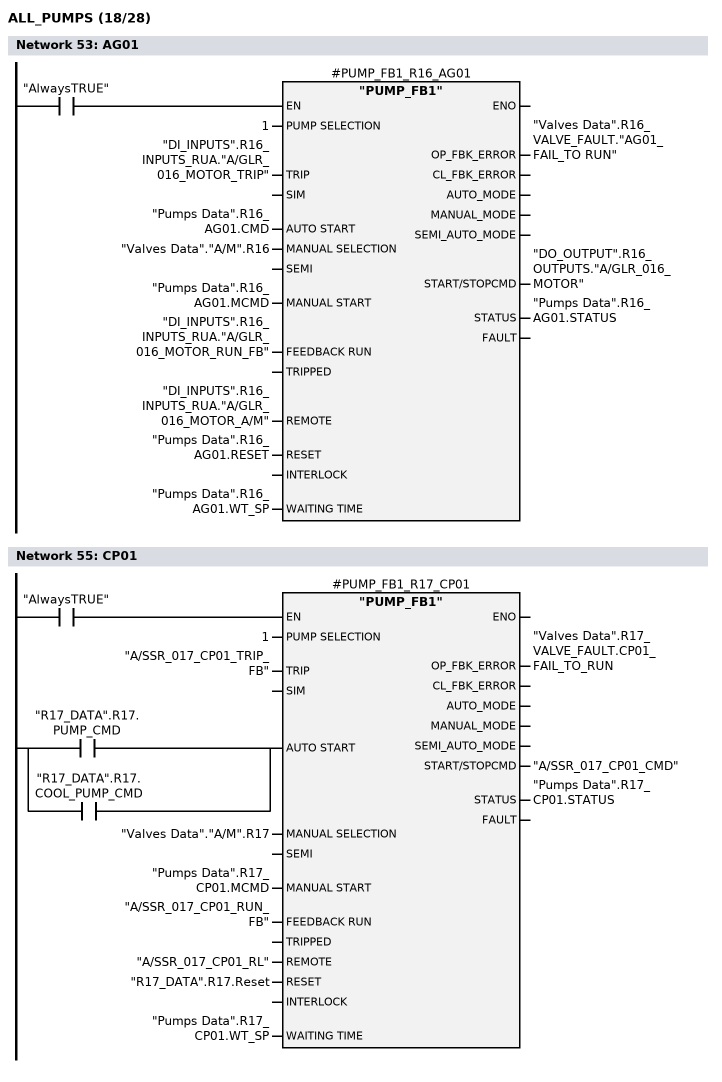
   RUNG wire#powerrail
      Contact( "AlwaysTRUE" )
      #PUMP_FB1_R16_AG01("PUMP SELECTION" := 1, TRIP := "DI_INPUTS".R16_INPUTS_RUA."A/GLR_016_MOTOR_TRIP", SIM :=, "AUTO START" := "Pumps Data".R16_AG01.CMD, "MANUAL SELECTION" := "Valves Data"."A/M".R16, SEMI :=, "MANUAL START" := "Pumps Data".R16_AG01.MCMD, "FEEDBACK RUN" := "DI_INPUTS".R16_INPUTS_RUA."A/GLR_016_MOTOR_RUN_FB", TRIPPED :=, REMOTE := "DI_INPUTS".R16_INPUTS_RUA."A/GLR_016_MOTOR_A/M", RESET := "Pumps Data".R16_AG01.RESET, INTERLOCK :=, "WAITING TIME" := "Pumps Data".R16_AG01.WT_SP, OP_FBK_ERROR => "Valves Data".R16_VALVE_FAULT."AG01_FAIL_TO RUN", CL_FBK_ERROR =>, AUTO_MODE =>, MANUAL_MODE =>, SEMI_AUTO_MODE =>, "START/STOPCMD" => "DO_OUTPUT".R16_OUTPUTS."A/GLR_016_MOTOR", STATUS => "Pumps Data".R16_AG01.STATUS, FAULT =>)
   END_RUNG
   // the same network as SCL:
   IF "AlwaysTRUE" THEN
       #PUMP_FB1_R16_AG01("PUMP SELECTION" := 1,   // "PUMP_FB1"
                          TRIP := "DI_INPUTS".R16_INPUTS_RUA."A/GLR_016_MOTOR_TRIP",
                          "AUTO START" := "Pumps Data".R16_AG01.CMD,
                          "MANUAL SELECTION" := "Valves Data"."A/M".R16,
                          "MANUAL START" := "Pumps Data".R16_AG01.MCMD,
                          "FEEDBACK RUN" := "DI_INPUTS".R16_INPUTS_RUA."A/GLR_016_MOTOR_RUN_FB",
                          REMOTE := "DI_INPUTS".R16_INPUTS_RUA."A/GLR_016_MOTOR_A/M",
                          RESET := "Pumps Data".R16_AG01.RESET,
                          "WAITING TIME" := "Pumps Data".R16_AG01.WT_SP,
                          OP_FBK_ERROR => "Valves Data".R16_VALVE_FAULT."AG01_FAIL_TO RUN",
                          "START/STOPCMD" => "DO_OUTPUT".R16_OUTPUTS."A/GLR_016_MOTOR",
                          STATUS => "Pumps Data".R16_AG01.STATUS);
   END_IF;
END_REGION

REGION Network 54: ***R17****
END_REGION

REGION Network 55: CP01
   RUNG wire#powerrail
      Contact( "AlwaysTRUE" )
      #PUMP_FB1_R17_CP01("AUTO START" := wire#w1, "PUMP SELECTION" := 1, TRIP := "A/SSR_017_CP01_TRIP_FB", SIM :=, "MANUAL SELECTION" := "Valves Data"."A/M".R17, SEMI :=, "MANUAL START" := "Pumps Data".R17_CP01.MCMD, "FEEDBACK RUN" := "A/SSR_017_CP01_RUN_FB", TRIPPED :=, REMOTE := "A/SSR_017_CP01_RL", RESET := "R17_DATA".R17.Reset, INTERLOCK :=, "WAITING TIME" := "Pumps Data".R17_CP01.WT_SP, OP_FBK_ERROR => "Valves Data".R17_VALVE_FAULT.CP01_FAIL_TO_RUN, CL_FBK_ERROR =>, AUTO_MODE =>, MANUAL_MODE =>, SEMI_AUTO_MODE =>, "START/STOPCMD" => "A/SSR_017_CP01_CMD", STATUS => "Pumps Data".R17_CP01.STATUS, FAULT =>)
   END_RUNG
   RUNG wire#powerrail
      Contact( "R17_DATA".R17.PUMP_CMD )
   END_RUNG wire#w1
   RUNG wire#powerrail
      Contact( "R17_DATA".R17.COOL_PUMP_CMD )
   END_RUNG wire#w1
   // the same network as SCL:
   IF "AlwaysTRUE" THEN
       #PUMP_FB1_R17_CP01("PUMP SELECTION" := 1,   // "PUMP_FB1"
                          TRIP := "A/SSR_017_CP01_TRIP_FB",
                          "AUTO START" := "R17_DATA".R17.PUMP_CMD OR "R17_DATA".R17.COOL_PUMP_CMD,
                          "MANUAL SELECTION" := "Valves Data"."A/M".R17,
                          "MANUAL START" := "Pumps Data".R17_CP01.MCMD,
                          "FEEDBACK RUN" := "A/SSR_017_CP01_RUN_FB",
                          REMOTE := "A/SSR_017_CP01_RL",
                          RESET := "R17_DATA".R17.Reset,
                          "WAITING TIME" := "Pumps Data".R17_CP01.WT_SP,
                          OP_FBK_ERROR => "Valves Data".R17_VALVE_FAULT.CP01_FAIL_TO_RUN,
                          "START/STOPCMD" => "A/SSR_017_CP01_CMD",
                          STATUS => "Pumps Data".R17_CP01.STATUS);
   END_IF;
END_REGION

REGION Network 56: AG01
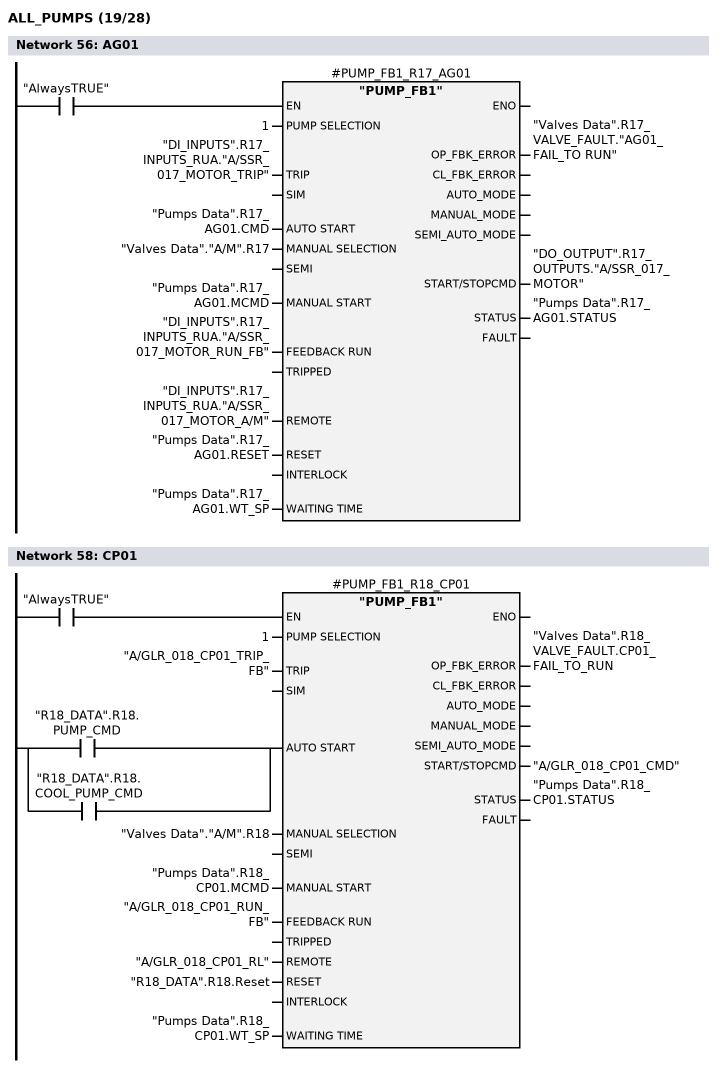
   RUNG wire#powerrail
      Contact( "AlwaysTRUE" )
      #PUMP_FB1_R17_AG01("PUMP SELECTION" := 1, TRIP := "DI_INPUTS".R17_INPUTS_RUA."A/SSR_017_MOTOR_TRIP", SIM :=, "AUTO START" := "Pumps Data".R17_AG01.CMD, "MANUAL SELECTION" := "Valves Data"."A/M".R17, SEMI :=, "MANUAL START" := "Pumps Data".R17_AG01.MCMD, "FEEDBACK RUN" := "DI_INPUTS".R17_INPUTS_RUA."A/SSR_017_MOTOR_RUN_FB", TRIPPED :=, REMOTE := "DI_INPUTS".R17_INPUTS_RUA."A/SSR_017_MOTOR_A/M", RESET := "Pumps Data".R17_AG01.RESET, INTERLOCK :=, "WAITING TIME" := "Pumps Data".R17_AG01.WT_SP, OP_FBK_ERROR => "Valves Data".R17_VALVE_FAULT."AG01_FAIL_TO RUN", CL_FBK_ERROR =>, AUTO_MODE =>, MANUAL_MODE =>, SEMI_AUTO_MODE =>, "START/STOPCMD" => "DO_OUTPUT".R17_OUTPUTS."A/SSR_017_MOTOR", STATUS => "Pumps Data".R17_AG01.STATUS, FAULT =>)
   END_RUNG
   // the same network as SCL:
   IF "AlwaysTRUE" THEN
       #PUMP_FB1_R17_AG01("PUMP SELECTION" := 1,   // "PUMP_FB1"
                          TRIP := "DI_INPUTS".R17_INPUTS_RUA."A/SSR_017_MOTOR_TRIP",
                          "AUTO START" := "Pumps Data".R17_AG01.CMD,
                          "MANUAL SELECTION" := "Valves Data"."A/M".R17,
                          "MANUAL START" := "Pumps Data".R17_AG01.MCMD,
                          "FEEDBACK RUN" := "DI_INPUTS".R17_INPUTS_RUA."A/SSR_017_MOTOR_RUN_FB",
                          REMOTE := "DI_INPUTS".R17_INPUTS_RUA."A/SSR_017_MOTOR_A/M",
                          RESET := "Pumps Data".R17_AG01.RESET,
                          "WAITING TIME" := "Pumps Data".R17_AG01.WT_SP,
                          OP_FBK_ERROR => "Valves Data".R17_VALVE_FAULT."AG01_FAIL_TO RUN",
                          "START/STOPCMD" => "DO_OUTPUT".R17_OUTPUTS."A/SSR_017_MOTOR",
                          STATUS => "Pumps Data".R17_AG01.STATUS);
   END_IF;
END_REGION

REGION Network 57: ***R18****
END_REGION

REGION Network 58: CP01
   RUNG wire#powerrail
      Contact( "AlwaysTRUE" )
      #PUMP_FB1_R18_CP01("AUTO START" := wire#w1, "PUMP SELECTION" := 1, TRIP := "A/GLR_018_CP01_TRIP_FB", SIM :=, "MANUAL SELECTION" := "Valves Data"."A/M".R18, SEMI :=, "MANUAL START" := "Pumps Data".R18_CP01.MCMD, "FEEDBACK RUN" := "A/GLR_018_CP01_RUN_FB", TRIPPED :=, REMOTE := "A/GLR_018_CP01_RL", RESET := "R18_DATA".R18.Reset, INTERLOCK :=, "WAITING TIME" := "Pumps Data".R18_CP01.WT_SP, OP_FBK_ERROR => "Valves Data".R18_VALVE_FAULT.CP01_FAIL_TO_RUN, CL_FBK_ERROR =>, AUTO_MODE =>, MANUAL_MODE =>, SEMI_AUTO_MODE =>, "START/STOPCMD" => "A/GLR_018_CP01_CMD", STATUS => "Pumps Data".R18_CP01.STATUS, FAULT =>)
   END_RUNG
   RUNG wire#powerrail
      Contact( "R18_DATA".R18.PUMP_CMD )
   END_RUNG wire#w1
   RUNG wire#powerrail
      Contact( "R18_DATA".R18.COOL_PUMP_CMD )
   END_RUNG wire#w1
   // the same network as SCL:
   IF "AlwaysTRUE" THEN
       #PUMP_FB1_R18_CP01("PUMP SELECTION" := 1,   // "PUMP_FB1"
                          TRIP := "A/GLR_018_CP01_TRIP_FB",
                          "AUTO START" := "R18_DATA".R18.PUMP_CMD OR "R18_DATA".R18.COOL_PUMP_CMD,
                          "MANUAL SELECTION" := "Valves Data"."A/M".R18,
                          "MANUAL START" := "Pumps Data".R18_CP01.MCMD,
                          "FEEDBACK RUN" := "A/GLR_018_CP01_RUN_FB",
                          REMOTE := "A/GLR_018_CP01_RL",
                          RESET := "R18_DATA".R18.Reset,
                          "WAITING TIME" := "Pumps Data".R18_CP01.WT_SP,
                          OP_FBK_ERROR => "Valves Data".R18_VALVE_FAULT.CP01_FAIL_TO_RUN,
                          "START/STOPCMD" => "A/GLR_018_CP01_CMD",
                          STATUS => "Pumps Data".R18_CP01.STATUS);
   END_IF;
END_REGION

REGION Network 59: AG01
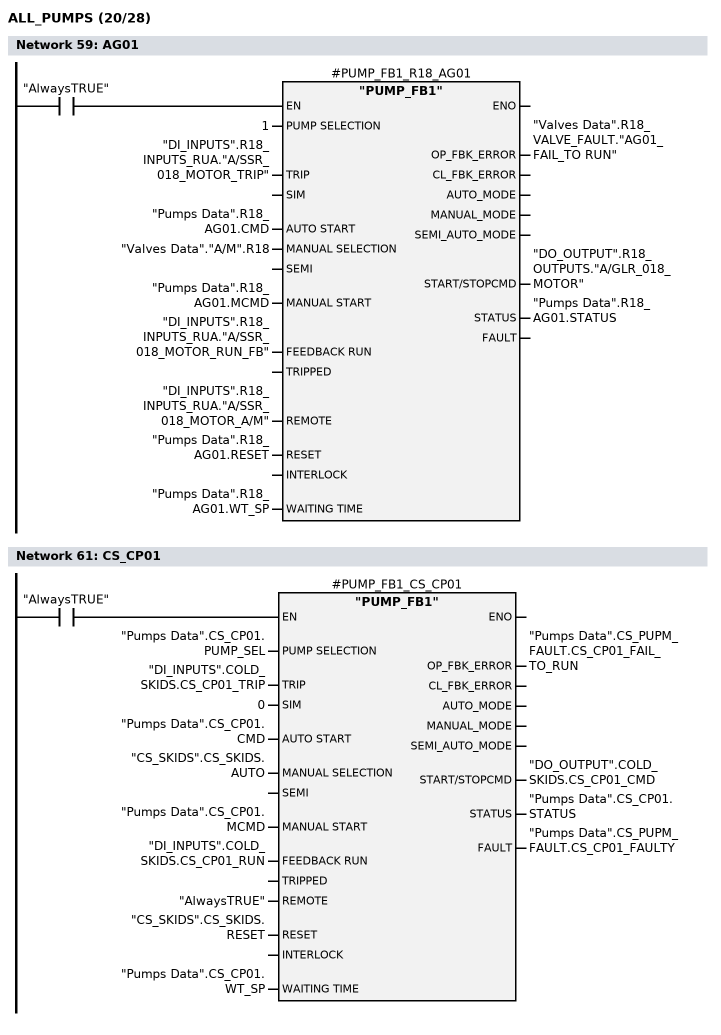
   RUNG wire#powerrail
      Contact( "AlwaysTRUE" )
      #PUMP_FB1_R18_AG01("PUMP SELECTION" := 1, TRIP := "DI_INPUTS".R18_INPUTS_RUA."A/SSR_018_MOTOR_TRIP", SIM :=, "AUTO START" := "Pumps Data".R18_AG01.CMD, "MANUAL SELECTION" := "Valves Data"."A/M".R18, SEMI :=, "MANUAL START" := "Pumps Data".R18_AG01.MCMD, "FEEDBACK RUN" := "DI_INPUTS".R18_INPUTS_RUA."A/SSR_018_MOTOR_RUN_FB", TRIPPED :=, REMOTE := "DI_INPUTS".R18_INPUTS_RUA."A/SSR_018_MOTOR_A/M", RESET := "Pumps Data".R18_AG01.RESET, INTERLOCK :=, "WAITING TIME" := "Pumps Data".R18_AG01.WT_SP, OP_FBK_ERROR => "Valves Data".R18_VALVE_FAULT."AG01_FAIL_TO RUN", CL_FBK_ERROR =>, AUTO_MODE =>, MANUAL_MODE =>, SEMI_AUTO_MODE =>, "START/STOPCMD" => "DO_OUTPUT".R18_OUTPUTS."A/GLR_018_MOTOR", STATUS => "Pumps Data".R18_AG01.STATUS, FAULT =>)
   END_RUNG
   // the same network as SCL:
   IF "AlwaysTRUE" THEN
       #PUMP_FB1_R18_AG01("PUMP SELECTION" := 1,   // "PUMP_FB1"
                          TRIP := "DI_INPUTS".R18_INPUTS_RUA."A/SSR_018_MOTOR_TRIP",
                          "AUTO START" := "Pumps Data".R18_AG01.CMD,
                          "MANUAL SELECTION" := "Valves Data"."A/M".R18,
                          "MANUAL START" := "Pumps Data".R18_AG01.MCMD,
                          "FEEDBACK RUN" := "DI_INPUTS".R18_INPUTS_RUA."A/SSR_018_MOTOR_RUN_FB",
                          REMOTE := "DI_INPUTS".R18_INPUTS_RUA."A/SSR_018_MOTOR_A/M",
                          RESET := "Pumps Data".R18_AG01.RESET,
                          "WAITING TIME" := "Pumps Data".R18_AG01.WT_SP,
                          OP_FBK_ERROR => "Valves Data".R18_VALVE_FAULT."AG01_FAIL_TO RUN",
                          "START/STOPCMD" => "DO_OUTPUT".R18_OUTPUTS."A/GLR_018_MOTOR",
                          STATUS => "Pumps Data".R18_AG01.STATUS);
   END_IF;
END_REGION

REGION Network 60: ****CS_SKIDS****
END_REGION

REGION Network 61: CS_CP01
   RUNG wire#powerrail
      Contact( "AlwaysTRUE" )
      #PUMP_FB1_CS_CP01("PUMP SELECTION" := "Pumps Data".CS_CP01.PUMP_SEL, TRIP := "DI_INPUTS".COLD_SKIDS.CS_CP01_TRIP, SIM := 0, "AUTO START" := "Pumps Data".CS_CP01.CMD, "MANUAL SELECTION" := "CS_SKIDS".CS_SKIDS.AUTO, SEMI :=, "MANUAL START" := "Pumps Data".CS_CP01.MCMD, "FEEDBACK RUN" := "DI_INPUTS".COLD_SKIDS.CS_CP01_RUN, TRIPPED :=, REMOTE := "AlwaysTRUE", RESET := "CS_SKIDS".CS_SKIDS.RESET, INTERLOCK :=, "WAITING TIME" := "Pumps Data".CS_CP01.WT_SP, OP_FBK_ERROR => "Pumps Data".CS_PUPM_FAULT.CS_CP01_FAIL_TO_RUN, CL_FBK_ERROR =>, AUTO_MODE =>, MANUAL_MODE =>, SEMI_AUTO_MODE =>, "START/STOPCMD" => "DO_OUTPUT".COLD_SKIDS.CS_CP01_CMD, STATUS => "Pumps Data".CS_CP01.STATUS, FAULT => "Pumps Data".CS_PUPM_FAULT.CS_CP01_FAULTY)
   END_RUNG
   // the same network as SCL:
   IF "AlwaysTRUE" THEN
       #PUMP_FB1_CS_CP01("PUMP SELECTION" := "Pumps Data".CS_CP01.PUMP_SEL,   // "PUMP_FB1"
                         TRIP := "DI_INPUTS".COLD_SKIDS.CS_CP01_TRIP,
                         SIM := 0,
                         "AUTO START" := "Pumps Data".CS_CP01.CMD,
                         "MANUAL SELECTION" := "CS_SKIDS".CS_SKIDS.AUTO,
                         "MANUAL START" := "Pumps Data".CS_CP01.MCMD,
                         "FEEDBACK RUN" := "DI_INPUTS".COLD_SKIDS.CS_CP01_RUN,
                         REMOTE := "AlwaysTRUE",
                         RESET := "CS_SKIDS".CS_SKIDS.RESET,
                         "WAITING TIME" := "Pumps Data".CS_CP01.WT_SP,
                         OP_FBK_ERROR => "Pumps Data".CS_PUPM_FAULT.CS_CP01_FAIL_TO_RUN,
                         "START/STOPCMD" => "DO_OUTPUT".COLD_SKIDS.CS_CP01_CMD,
                         STATUS => "Pumps Data".CS_CP01.STATUS,
                         FAULT => "Pumps Data".CS_PUPM_FAULT.CS_CP01_FAULTY);
   END_IF;
END_REGION

REGION Network 62: CS_CP02
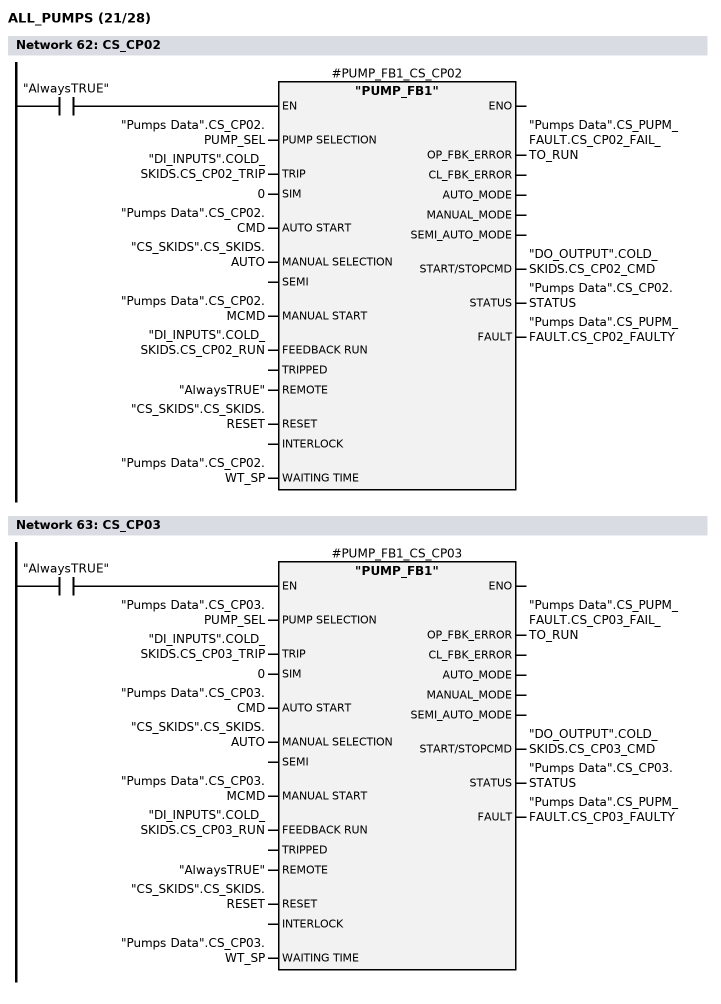
   RUNG wire#powerrail
      Contact( "AlwaysTRUE" )
      #PUMP_FB1_CS_CP02("PUMP SELECTION" := "Pumps Data".CS_CP02.PUMP_SEL, TRIP := "DI_INPUTS".COLD_SKIDS.CS_CP02_TRIP, SIM := 0, "AUTO START" := "Pumps Data".CS_CP02.CMD, "MANUAL SELECTION" := "CS_SKIDS".CS_SKIDS.AUTO, SEMI :=, "MANUAL START" := "Pumps Data".CS_CP02.MCMD, "FEEDBACK RUN" := "DI_INPUTS".COLD_SKIDS.CS_CP02_RUN, TRIPPED :=, REMOTE := "AlwaysTRUE", RESET := "CS_SKIDS".CS_SKIDS.RESET, INTERLOCK :=, "WAITING TIME" := "Pumps Data".CS_CP02.WT_SP, OP_FBK_ERROR => "Pumps Data".CS_PUPM_FAULT.CS_CP02_FAIL_TO_RUN, CL_FBK_ERROR =>, AUTO_MODE =>, MANUAL_MODE =>, SEMI_AUTO_MODE =>, "START/STOPCMD" => "DO_OUTPUT".COLD_SKIDS.CS_CP02_CMD, STATUS => "Pumps Data".CS_CP02.STATUS, FAULT => "Pumps Data".CS_PUPM_FAULT.CS_CP02_FAULTY)
   END_RUNG
   // the same network as SCL:
   IF "AlwaysTRUE" THEN
       #PUMP_FB1_CS_CP02("PUMP SELECTION" := "Pumps Data".CS_CP02.PUMP_SEL,   // "PUMP_FB1"
                         TRIP := "DI_INPUTS".COLD_SKIDS.CS_CP02_TRIP,
                         SIM := 0,
                         "AUTO START" := "Pumps Data".CS_CP02.CMD,
                         "MANUAL SELECTION" := "CS_SKIDS".CS_SKIDS.AUTO,
                         "MANUAL START" := "Pumps Data".CS_CP02.MCMD,
                         "FEEDBACK RUN" := "DI_INPUTS".COLD_SKIDS.CS_CP02_RUN,
                         REMOTE := "AlwaysTRUE",
                         RESET := "CS_SKIDS".CS_SKIDS.RESET,
                         "WAITING TIME" := "Pumps Data".CS_CP02.WT_SP,
                         OP_FBK_ERROR => "Pumps Data".CS_PUPM_FAULT.CS_CP02_FAIL_TO_RUN,
                         "START/STOPCMD" => "DO_OUTPUT".COLD_SKIDS.CS_CP02_CMD,
                         STATUS => "Pumps Data".CS_CP02.STATUS,
                         FAULT => "Pumps Data".CS_PUPM_FAULT.CS_CP02_FAULTY);
   END_IF;
END_REGION

REGION Network 63: CS_CP03
   RUNG wire#powerrail
      Contact( "AlwaysTRUE" )
      #PUMP_FB1_CS_CP03("PUMP SELECTION" := "Pumps Data".CS_CP03.PUMP_SEL, TRIP := "DI_INPUTS".COLD_SKIDS.CS_CP03_TRIP, SIM := 0, "AUTO START" := "Pumps Data".CS_CP03.CMD, "MANUAL SELECTION" := "CS_SKIDS".CS_SKIDS.AUTO, SEMI :=, "MANUAL START" := "Pumps Data".CS_CP03.MCMD, "FEEDBACK RUN" := "DI_INPUTS".COLD_SKIDS.CS_CP03_RUN, TRIPPED :=, REMOTE := "AlwaysTRUE", RESET := "CS_SKIDS".CS_SKIDS.RESET, INTERLOCK :=, "WAITING TIME" := "Pumps Data".CS_CP03.WT_SP, OP_FBK_ERROR => "Pumps Data".CS_PUPM_FAULT.CS_CP03_FAIL_TO_RUN, CL_FBK_ERROR =>, AUTO_MODE =>, MANUAL_MODE =>, SEMI_AUTO_MODE =>, "START/STOPCMD" => "DO_OUTPUT".COLD_SKIDS.CS_CP03_CMD, STATUS => "Pumps Data".CS_CP03.STATUS, FAULT => "Pumps Data".CS_PUPM_FAULT.CS_CP03_FAULTY)
   END_RUNG
   // the same network as SCL:
   IF "AlwaysTRUE" THEN
       #PUMP_FB1_CS_CP03("PUMP SELECTION" := "Pumps Data".CS_CP03.PUMP_SEL,   // "PUMP_FB1"
                         TRIP := "DI_INPUTS".COLD_SKIDS.CS_CP03_TRIP,
                         SIM := 0,
                         "AUTO START" := "Pumps Data".CS_CP03.CMD,
                         "MANUAL SELECTION" := "CS_SKIDS".CS_SKIDS.AUTO,
                         "MANUAL START" := "Pumps Data".CS_CP03.MCMD,
                         "FEEDBACK RUN" := "DI_INPUTS".COLD_SKIDS.CS_CP03_RUN,
                         REMOTE := "AlwaysTRUE",
                         RESET := "CS_SKIDS".CS_SKIDS.RESET,
                         "WAITING TIME" := "Pumps Data".CS_CP03.WT_SP,
                         OP_FBK_ERROR => "Pumps Data".CS_PUPM_FAULT.CS_CP03_FAIL_TO_RUN,
                         "START/STOPCMD" => "DO_OUTPUT".COLD_SKIDS.CS_CP03_CMD,
                         STATUS => "Pumps Data".CS_CP03.STATUS,
                         FAULT => "Pumps Data".CS_PUPM_FAULT.CS_CP03_FAULTY);
   END_IF;
END_REGION

REGION Network 64: ****UCHS_SKIDS****
END_REGION

REGION Network 65: UCHS_CP01
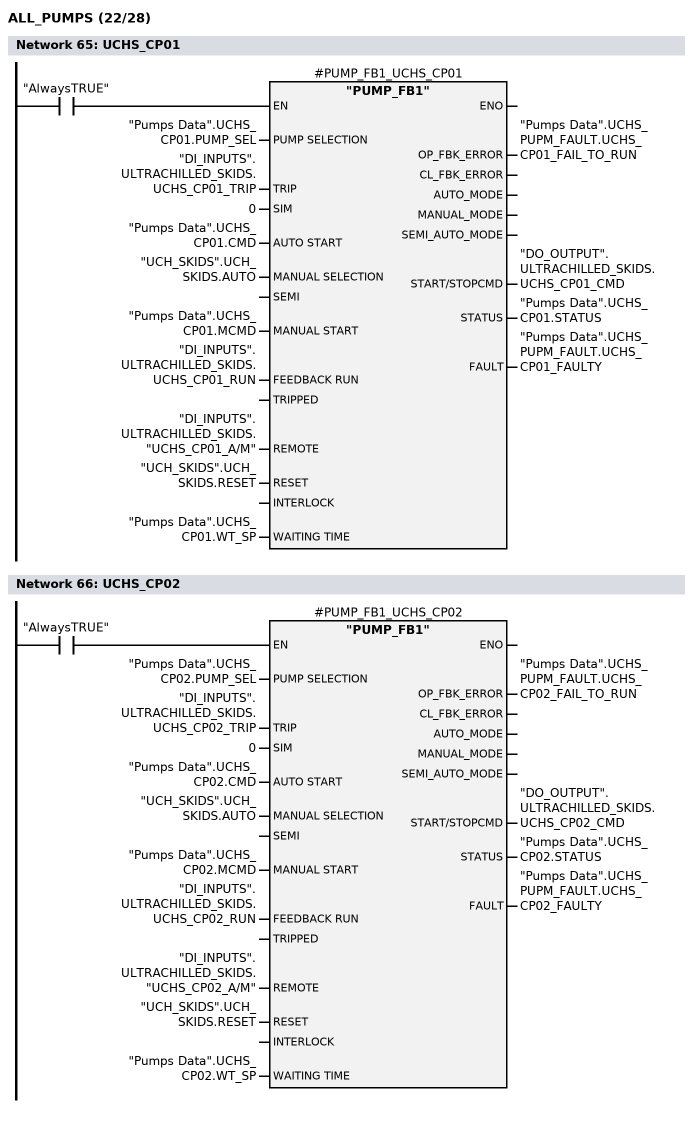
   RUNG wire#powerrail
      Contact( "AlwaysTRUE" )
      #PUMP_FB1_UCHS_CP01("PUMP SELECTION" := "Pumps Data".UCHS_CP01.PUMP_SEL, TRIP := "DI_INPUTS".ULTRACHILLED_SKIDS.UCHS_CP01_TRIP, SIM := 0, "AUTO START" := "Pumps Data".UCHS_CP01.CMD, "MANUAL SELECTION" := "UCH_SKIDS".UCH_SKIDS.AUTO, SEMI :=, "MANUAL START" := "Pumps Data".UCHS_CP01.MCMD, "FEEDBACK RUN" := "DI_INPUTS".ULTRACHILLED_SKIDS.UCHS_CP01_RUN, TRIPPED :=, REMOTE := "DI_INPUTS".ULTRACHILLED_SKIDS."UCHS_CP01_A/M", RESET := "UCH_SKIDS".UCH_SKIDS.RESET, INTERLOCK :=, "WAITING TIME" := "Pumps Data".UCHS_CP01.WT_SP, OP_FBK_ERROR => "Pumps Data".UCHS_PUPM_FAULT.UCHS_CP01_FAIL_TO_RUN, CL_FBK_ERROR =>, AUTO_MODE =>, MANUAL_MODE =>, SEMI_AUTO_MODE =>, "START/STOPCMD" => "DO_OUTPUT".ULTRACHILLED_SKIDS.UCHS_CP01_CMD, STATUS => "Pumps Data".UCHS_CP01.STATUS, FAULT => "Pumps Data".UCHS_PUPM_FAULT.UCHS_CP01_FAULTY)
   END_RUNG
   // the same network as SCL:
   IF "AlwaysTRUE" THEN
       #PUMP_FB1_UCHS_CP01("PUMP SELECTION" := "Pumps Data".UCHS_CP01.PUMP_SEL,   // "PUMP_FB1"
                           TRIP := "DI_INPUTS".ULTRACHILLED_SKIDS.UCHS_CP01_TRIP,
                           SIM := 0,
                           "AUTO START" := "Pumps Data".UCHS_CP01.CMD,
                           "MANUAL SELECTION" := "UCH_SKIDS".UCH_SKIDS.AUTO,
                           "MANUAL START" := "Pumps Data".UCHS_CP01.MCMD,
                           "FEEDBACK RUN" := "DI_INPUTS".ULTRACHILLED_SKIDS.UCHS_CP01_RUN,
                           REMOTE := "DI_INPUTS".ULTRACHILLED_SKIDS."UCHS_CP01_A/M",
                           RESET := "UCH_SKIDS".UCH_SKIDS.RESET,
                           "WAITING TIME" := "Pumps Data".UCHS_CP01.WT_SP,
                           OP_FBK_ERROR => "Pumps Data".UCHS_PUPM_FAULT.UCHS_CP01_FAIL_TO_RUN,
                           "START/STOPCMD" => "DO_OUTPUT".ULTRACHILLED_SKIDS.UCHS_CP01_CMD,
                           STATUS => "Pumps Data".UCHS_CP01.STATUS,
                           FAULT => "Pumps Data".UCHS_PUPM_FAULT.UCHS_CP01_FAULTY);
   END_IF;
END_REGION

REGION Network 66: UCHS_CP02
   RUNG wire#powerrail
      Contact( "AlwaysTRUE" )
      #PUMP_FB1_UCHS_CP02("PUMP SELECTION" := "Pumps Data".UCHS_CP02.PUMP_SEL, TRIP := "DI_INPUTS".ULTRACHILLED_SKIDS.UCHS_CP02_TRIP, SIM := 0, "AUTO START" := "Pumps Data".UCHS_CP02.CMD, "MANUAL SELECTION" := "UCH_SKIDS".UCH_SKIDS.AUTO, SEMI :=, "MANUAL START" := "Pumps Data".UCHS_CP02.MCMD, "FEEDBACK RUN" := "DI_INPUTS".ULTRACHILLED_SKIDS.UCHS_CP02_RUN, TRIPPED :=, REMOTE := "DI_INPUTS".ULTRACHILLED_SKIDS."UCHS_CP02_A/M", RESET := "UCH_SKIDS".UCH_SKIDS.RESET, INTERLOCK :=, "WAITING TIME" := "Pumps Data".UCHS_CP02.WT_SP, OP_FBK_ERROR => "Pumps Data".UCHS_PUPM_FAULT.UCHS_CP02_FAIL_TO_RUN, CL_FBK_ERROR =>, AUTO_MODE =>, MANUAL_MODE =>, SEMI_AUTO_MODE =>, "START/STOPCMD" => "DO_OUTPUT".ULTRACHILLED_SKIDS.UCHS_CP02_CMD, STATUS => "Pumps Data".UCHS_CP02.STATUS, FAULT => "Pumps Data".UCHS_PUPM_FAULT.UCHS_CP02_FAULTY)
   END_RUNG
   // the same network as SCL:
   IF "AlwaysTRUE" THEN
       #PUMP_FB1_UCHS_CP02("PUMP SELECTION" := "Pumps Data".UCHS_CP02.PUMP_SEL,   // "PUMP_FB1"
                           TRIP := "DI_INPUTS".ULTRACHILLED_SKIDS.UCHS_CP02_TRIP,
                           SIM := 0,
                           "AUTO START" := "Pumps Data".UCHS_CP02.CMD,
                           "MANUAL SELECTION" := "UCH_SKIDS".UCH_SKIDS.AUTO,
                           "MANUAL START" := "Pumps Data".UCHS_CP02.MCMD,
                           "FEEDBACK RUN" := "DI_INPUTS".ULTRACHILLED_SKIDS.UCHS_CP02_RUN,
                           REMOTE := "DI_INPUTS".ULTRACHILLED_SKIDS."UCHS_CP02_A/M",
                           RESET := "UCH_SKIDS".UCH_SKIDS.RESET,
                           "WAITING TIME" := "Pumps Data".UCHS_CP02.WT_SP,
                           OP_FBK_ERROR => "Pumps Data".UCHS_PUPM_FAULT.UCHS_CP02_FAIL_TO_RUN,
                           "START/STOPCMD" => "DO_OUTPUT".ULTRACHILLED_SKIDS.UCHS_CP02_CMD,
                           STATUS => "Pumps Data".UCHS_CP02.STATUS,
                           FAULT => "Pumps Data".UCHS_PUPM_FAULT.UCHS_CP02_FAULTY);
   END_IF;
END_REGION

REGION Network 67: ****HS_SKIDS****
END_REGION

REGION Network 68: HS_CP01
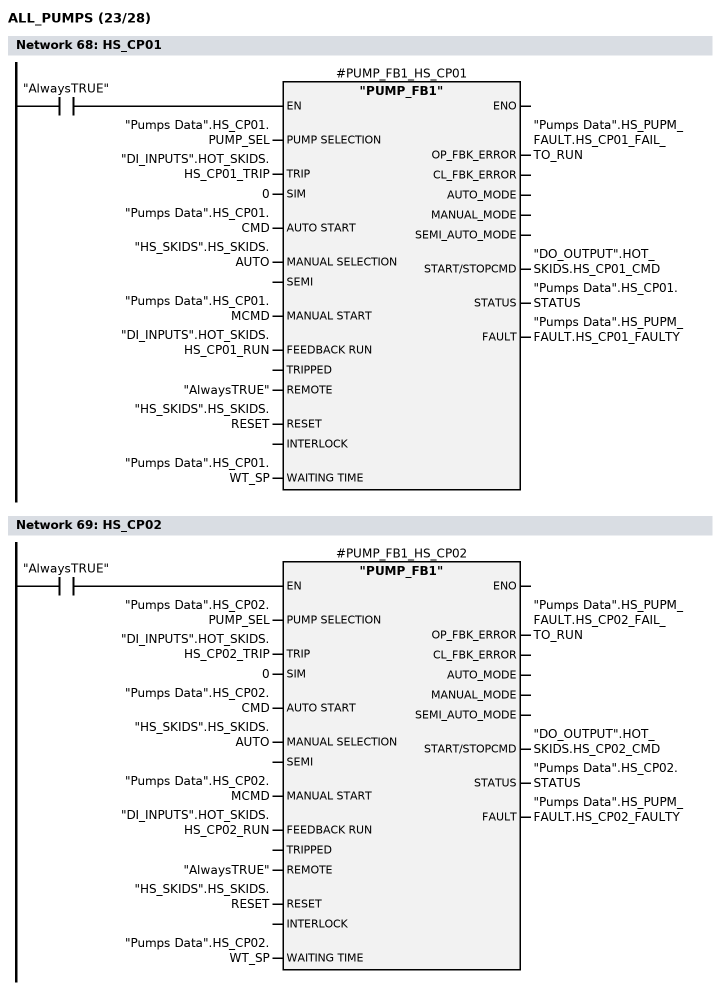
   RUNG wire#powerrail
      Contact( "AlwaysTRUE" )
      #PUMP_FB1_HS_CP01("PUMP SELECTION" := "Pumps Data".HS_CP01.PUMP_SEL, TRIP := "DI_INPUTS".HOT_SKIDS.HS_CP01_TRIP, SIM := 0, "AUTO START" := "Pumps Data".HS_CP01.CMD, "MANUAL SELECTION" := "HS_SKIDS".HS_SKIDS.AUTO, SEMI :=, "MANUAL START" := "Pumps Data".HS_CP01.MCMD, "FEEDBACK RUN" := "DI_INPUTS".HOT_SKIDS.HS_CP01_RUN, TRIPPED :=, REMOTE := "AlwaysTRUE", RESET := "HS_SKIDS".HS_SKIDS.RESET, INTERLOCK :=, "WAITING TIME" := "Pumps Data".HS_CP01.WT_SP, OP_FBK_ERROR => "Pumps Data".HS_PUPM_FAULT.HS_CP01_FAIL_TO_RUN, CL_FBK_ERROR =>, AUTO_MODE =>, MANUAL_MODE =>, SEMI_AUTO_MODE =>, "START/STOPCMD" => "DO_OUTPUT".HOT_SKIDS.HS_CP01_CMD, STATUS => "Pumps Data".HS_CP01.STATUS, FAULT => "Pumps Data".HS_PUPM_FAULT.HS_CP01_FAULTY)
   END_RUNG
   // the same network as SCL:
   IF "AlwaysTRUE" THEN
       #PUMP_FB1_HS_CP01("PUMP SELECTION" := "Pumps Data".HS_CP01.PUMP_SEL,   // "PUMP_FB1"
                         TRIP := "DI_INPUTS".HOT_SKIDS.HS_CP01_TRIP,
                         SIM := 0,
                         "AUTO START" := "Pumps Data".HS_CP01.CMD,
                         "MANUAL SELECTION" := "HS_SKIDS".HS_SKIDS.AUTO,
                         "MANUAL START" := "Pumps Data".HS_CP01.MCMD,
                         "FEEDBACK RUN" := "DI_INPUTS".HOT_SKIDS.HS_CP01_RUN,
                         REMOTE := "AlwaysTRUE",
                         RESET := "HS_SKIDS".HS_SKIDS.RESET,
                         "WAITING TIME" := "Pumps Data".HS_CP01.WT_SP,
                         OP_FBK_ERROR => "Pumps Data".HS_PUPM_FAULT.HS_CP01_FAIL_TO_RUN,
                         "START/STOPCMD" => "DO_OUTPUT".HOT_SKIDS.HS_CP01_CMD,
                         STATUS => "Pumps Data".HS_CP01.STATUS,
                         FAULT => "Pumps Data".HS_PUPM_FAULT.HS_CP01_FAULTY);
   END_IF;
END_REGION

REGION Network 69: HS_CP02
   RUNG wire#powerrail
      Contact( "AlwaysTRUE" )
      #PUMP_FB1_HS_CP02("PUMP SELECTION" := "Pumps Data".HS_CP02.PUMP_SEL, TRIP := "DI_INPUTS".HOT_SKIDS.HS_CP02_TRIP, SIM := 0, "AUTO START" := "Pumps Data".HS_CP02.CMD, "MANUAL SELECTION" := "HS_SKIDS".HS_SKIDS.AUTO, SEMI :=, "MANUAL START" := "Pumps Data".HS_CP02.MCMD, "FEEDBACK RUN" := "DI_INPUTS".HOT_SKIDS.HS_CP02_RUN, TRIPPED :=, REMOTE := "AlwaysTRUE", RESET := "HS_SKIDS".HS_SKIDS.RESET, INTERLOCK :=, "WAITING TIME" := "Pumps Data".HS_CP02.WT_SP, OP_FBK_ERROR => "Pumps Data".HS_PUPM_FAULT.HS_CP02_FAIL_TO_RUN, CL_FBK_ERROR =>, AUTO_MODE =>, MANUAL_MODE =>, SEMI_AUTO_MODE =>, "START/STOPCMD" => "DO_OUTPUT".HOT_SKIDS.HS_CP02_CMD, STATUS => "Pumps Data".HS_CP02.STATUS, FAULT => "Pumps Data".HS_PUPM_FAULT.HS_CP02_FAULTY)
   END_RUNG
   // the same network as SCL:
   IF "AlwaysTRUE" THEN
       #PUMP_FB1_HS_CP02("PUMP SELECTION" := "Pumps Data".HS_CP02.PUMP_SEL,   // "PUMP_FB1"
                         TRIP := "DI_INPUTS".HOT_SKIDS.HS_CP02_TRIP,
                         SIM := 0,
                         "AUTO START" := "Pumps Data".HS_CP02.CMD,
                         "MANUAL SELECTION" := "HS_SKIDS".HS_SKIDS.AUTO,
                         "MANUAL START" := "Pumps Data".HS_CP02.MCMD,
                         "FEEDBACK RUN" := "DI_INPUTS".HOT_SKIDS.HS_CP02_RUN,
                         REMOTE := "AlwaysTRUE",
                         RESET := "HS_SKIDS".HS_SKIDS.RESET,
                         "WAITING TIME" := "Pumps Data".HS_CP02.WT_SP,
                         OP_FBK_ERROR => "Pumps Data".HS_PUPM_FAULT.HS_CP02_FAIL_TO_RUN,
                         "START/STOPCMD" => "DO_OUTPUT".HOT_SKIDS.HS_CP02_CMD,
                         STATUS => "Pumps Data".HS_CP02.STATUS,
                         FAULT => "Pumps Data".HS_PUPM_FAULT.HS_CP02_FAULTY);
   END_IF;
END_REGION

REGION Network 70: HS_CP03
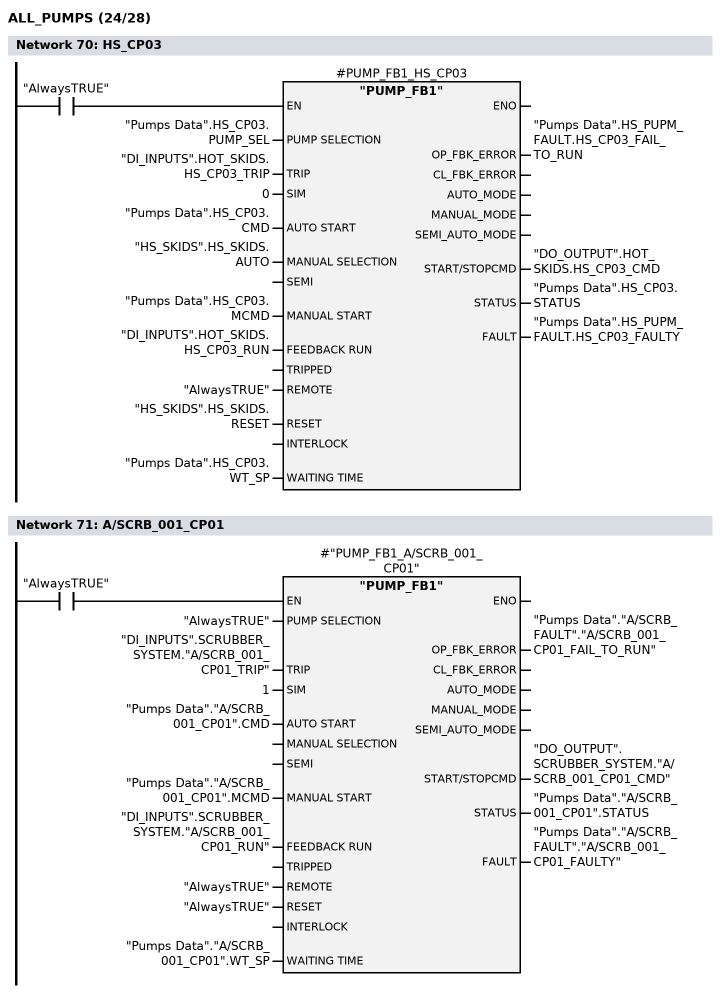
   RUNG wire#powerrail
      Contact( "AlwaysTRUE" )
      #PUMP_FB1_HS_CP03("PUMP SELECTION" := "Pumps Data".HS_CP03.PUMP_SEL, TRIP := "DI_INPUTS".HOT_SKIDS.HS_CP03_TRIP, SIM := 0, "AUTO START" := "Pumps Data".HS_CP03.CMD, "MANUAL SELECTION" := "HS_SKIDS".HS_SKIDS.AUTO, SEMI :=, "MANUAL START" := "Pumps Data".HS_CP03.MCMD, "FEEDBACK RUN" := "DI_INPUTS".HOT_SKIDS.HS_CP03_RUN, TRIPPED :=, REMOTE := "AlwaysTRUE", RESET := "HS_SKIDS".HS_SKIDS.RESET, INTERLOCK :=, "WAITING TIME" := "Pumps Data".HS_CP03.WT_SP, OP_FBK_ERROR => "Pumps Data".HS_PUPM_FAULT.HS_CP03_FAIL_TO_RUN, CL_FBK_ERROR =>, AUTO_MODE =>, MANUAL_MODE =>, SEMI_AUTO_MODE =>, "START/STOPCMD" => "DO_OUTPUT".HOT_SKIDS.HS_CP03_CMD, STATUS => "Pumps Data".HS_CP03.STATUS, FAULT => "Pumps Data".HS_PUPM_FAULT.HS_CP03_FAULTY)
   END_RUNG
   // the same network as SCL:
   IF "AlwaysTRUE" THEN
       #PUMP_FB1_HS_CP03("PUMP SELECTION" := "Pumps Data".HS_CP03.PUMP_SEL,   // "PUMP_FB1"
                         TRIP := "DI_INPUTS".HOT_SKIDS.HS_CP03_TRIP,
                         SIM := 0,
                         "AUTO START" := "Pumps Data".HS_CP03.CMD,
                         "MANUAL SELECTION" := "HS_SKIDS".HS_SKIDS.AUTO,
                         "MANUAL START" := "Pumps Data".HS_CP03.MCMD,
                         "FEEDBACK RUN" := "DI_INPUTS".HOT_SKIDS.HS_CP03_RUN,
                         REMOTE := "AlwaysTRUE",
                         RESET := "HS_SKIDS".HS_SKIDS.RESET,
                         "WAITING TIME" := "Pumps Data".HS_CP03.WT_SP,
                         OP_FBK_ERROR => "Pumps Data".HS_PUPM_FAULT.HS_CP03_FAIL_TO_RUN,
                         "START/STOPCMD" => "DO_OUTPUT".HOT_SKIDS.HS_CP03_CMD,
                         STATUS => "Pumps Data".HS_CP03.STATUS,
                         FAULT => "Pumps Data".HS_PUPM_FAULT.HS_CP03_FAULTY);
   END_IF;
END_REGION

REGION Network 71: A/SCRB_001_CP01
   RUNG wire#powerrail
      Contact( "AlwaysTRUE" )
      #"PUMP_FB1_A/SCRB_001_CP01"("PUMP SELECTION" := "AlwaysTRUE", TRIP := "DI_INPUTS".SCRUBBER_SYSTEM."A/SCRB_001_CP01_TRIP", SIM := 1, "AUTO START" := "Pumps Data"."A/SCRB_001_CP01".CMD, "MANUAL SELECTION" :=, SEMI :=, "MANUAL START" := "Pumps Data"."A/SCRB_001_CP01".MCMD, "FEEDBACK RUN" := "DI_INPUTS".SCRUBBER_SYSTEM."A/SCRB_001_CP01_RUN", TRIPPED :=, REMOTE := "AlwaysTRUE", RESET := "AlwaysTRUE", INTERLOCK :=, "WAITING TIME" := "Pumps Data"."A/SCRB_001_CP01".WT_SP, OP_FBK_ERROR => "Pumps Data"."A/SCRB_FAULT"."A/SCRB_001_CP01_FAIL_TO_RUN", CL_FBK_ERROR =>, AUTO_MODE =>, MANUAL_MODE =>, SEMI_AUTO_MODE =>, "START/STOPCMD" => "DO_OUTPUT".SCRUBBER_SYSTEM."A/SCRB_001_CP01_CMD", STATUS => "Pumps Data"."A/SCRB_001_CP01".STATUS, FAULT => "Pumps Data"."A/SCRB_FAULT"."A/SCRB_001_CP01_FAULTY")
   END_RUNG
   // the same network as SCL:
   IF "AlwaysTRUE" THEN
       #"PUMP_FB1_A/SCRB_001_CP01"("PUMP SELECTION" := "AlwaysTRUE",   // "PUMP_FB1"
                               TRIP := "DI_INPUTS".SCRUBBER_SYSTEM."A/SCRB_001_CP01_TRIP",
                               SIM := 1,
                               "AUTO START" := "Pumps Data"."A/SCRB_001_CP01".CMD,
                               "MANUAL START" := "Pumps Data"."A/SCRB_001_CP01".MCMD,
                               "FEEDBACK RUN" := "DI_INPUTS".SCRUBBER_SYSTEM."A/SCRB_001_CP01_RUN",
                               REMOTE := "AlwaysTRUE",
                               RESET := "AlwaysTRUE",
                               "WAITING TIME" := "Pumps Data"."A/SCRB_001_CP01".WT_SP,
                               OP_FBK_ERROR => "Pumps Data"."A/SCRB_FAULT"."A/SCRB_001_CP01_FAIL_TO_RUN",
                               "START/STOPCMD" => "DO_OUTPUT".SCRUBBER_SYSTEM."A/SCRB_001_CP01_CMD",
                               STATUS => "Pumps Data"."A/SCRB_001_CP01".STATUS,
                               FAULT => "Pumps Data"."A/SCRB_FAULT"."A/SCRB_001_CP01_FAULTY");
   END_IF;
END_REGION

REGION Network 72: A/SCRB_001_CP02
